(* Logix 5000 project; controller TFF vendor 1 type 14 code 107 rev 34.11; software revision 34.03; part 2 of 36 *)

        [3,10].HIHIAlarmONS := 1, [3,10].FeedPumpTag := 1, [3,10].Value := 4, [3,10].ValueHMI := 4, [3,10].PV := 20.567827, [3,10].HITimer.EN := 1, [3,10].HITimer.DN := 1, [3,10].HIHITimer.EN := 1, [3,10].HIHITimer.DN := 1, [3,10].EnableCfg := 1, [3,11].HIAlarm := 1, [3,11].HIHIAlarm := 1, [3,11].LOLODisable := 1, [3,11].LODisable := 1, [3,11].FeedPumpEnable := 1, [3,11].HIAlarmONS := 1, [3,11].HIHIAlarmONS := 1, [3,11].FeedPumpTag := 1, [3,11].Value := 4, [3,11].ValueHMI := 4, [3,11].PV := 25.7337, [3,11].HITimer.EN := 1, [3,11].HITimer.DN := 1, [3,11].HIHITimer.EN := 1, [3,11].HIHITimer.DN := 1, [3,11].EnableCfg := 1, [3,12].HIAlarm := 1, [3,12].HIHIAlarm := 1, [3,12].LOLODisable := 1, [3,12].LODisable := 1, [3,12].TransferPumpEnable := 1, [3,12].HIAlarmONS := 1, [3,12].HIHIAlarmONS := 1, [3,12].TransferPumpTag := 2, [3,12].Value := 4, [3,12].ValueHMI := 4, [3,12].PV := 28.0231, [3,12].HITimer.EN := 1, [3,12].HITimer.DN := 1, [3,12].HIHITimer.EN := 1, [3,12].HIHITimer.DN := 1, [3,12].EnableCfg := 1, [3,13].HIAlarm := 1, [3,13].HIHIAlarm := 1, [3,13].LOLODisable := 1, [3,13].LODisable := 1, [3,13].TransferPumpEnable := 1, [3,13].HIAlarmONS := 1, [3,13].HIHIAlarmONS := 1, [3,13].TransferPumpTag := 2, [3,13].Value := 4, [3,13].ValueHMI := 4, [3,13].PV := 21.08868, [3,13].HITimer.EN := 1, [3,13].HITimer.DN := 1, [3,13].HIHITimer.EN := 1, [3,13].HIHITimer.DN := 1, [3,13].EnableCfg := 1, [3,28].PV := -1.048729, [3,28].EnableCfg := 1,
        [3,29].HIAlarm := 1, [3,29].HIHIAlarm := 1, [3,29].HIAlarmONS := 1, [3,29].HIHIAlarmONS := 1, [3,29].Value := 4, [3,29].ValueHMI := 4, [3,29].PV := 100.96327, [3,29].HITimer.EN := 1, [3,29].HITimer.DN := 1, [3,29].HIHITimer.EN := 1, [3,29].HIHITimer.DN := 1, [3,29].EnableCfg := 1, [3,30].HIAlarm := 1, [3,30].HIHIAlarm := 1, [3,30].HIAlarmONS := 1, [3,30].HIHIAlarmONS := 1, [3,30].Value := 4, [3,30].ValueHMI := 4, [3,30].PV := 0.024414062, [3,30].HITimer.EN := 1, [3,30].HITimer.DN := 1, [3,30].HIHITimer.EN := 1, [3,30].HIHITimer.DN := 1, [3,30].EnableCfg := 1, [3,31].HIAlarm := 1, [3,31].HIHIAlarm := 1, [3,31].HIAlarmONS := 1, [3,31].HIHIAlarmONS := 1, [3,31].Value := 4, [3,31].ValueHMI := 4, [3,31].PV := 9.026997, [3,31].HITimer.EN := 1, [3,31].HITimer.DN := 1, [3,31].HIHITimer.EN := 1, [3,31].HIHITimer.DN := 1, [3,31].EnableCfg := 1, [3,40].LOLODisable := 1, [3,40].LODisable := 1, [3,40].FeedPumpEnable := 1, [3,40].TransferPumpEnable := 1, [3,40].FeedPumpTag := 1, [3,40].TransferPumpTag := 2, [3,40].PV := 48.590927, [3,40].EnableCfg := 1, [3,41].LOLODisable := 1, [3,41].LODisable := 1, [3,41].FeedPumpEnable := 1, [3,41].TransferPumpEnable := 1, [3,41].FeedPumpTag := 1, [3,41].TransferPumpTag := 2, [3,41].PV := 5830.911, [3,41].EnableCfg := 1, [3,42].LOLODisable := 1, [3,42].LODisable := 1, [3,42].FeedPumpEnable := 1, [3,42].FeedPumpTag := 1, [3,42].PV := 2468.1392, [3,42].EnableCfg := 1, [3,43].LOLODisable := 1, [3,43].LODisable := 1,
        [3,43].TransferPumpEnable := 1, [3,43].TransferPumpTag := 2, [3,43].PV := 3362.772, [3,43].EnableCfg := 1, [4,0].Override := 1, [4,0].LOLODisable := 1, [4,0].LODisable := 1, [4,0].LOLOAlarmONS := 1, [4,0].LOAlarmONS := 1, [4,0].HIAlarmONS := 1, [4,0].HIHIAlarmONS := 1, [4,0].HI := 100.0, [4,0].HIHI := 100.0, [4,0].PV := -2.4997964, [4,0].LOLOTimer.PRE := 2000, [4,0].LOLOTimerSP := 2, [4,0].LOTimer.PRE := 2000, [4,0].LOTimerSP := 2, [4,0].HITimer.PRE := 2000, [4,0].HITimerSP := 2, [4,0].HIHITimer.PRE := 2000, [4,0].HIHITimerSP := 2, [4,1].Override := 1, [4,1].LOLO := 20.0, [4,1].LO := 20.0, [4,1].HI := 50.0, [4,1].HIHI := 50.0, [4,1].PV := -12.498303, [4,1].LOLOTimer.PRE := 2000, [4,1].LOLOTimerSP := 2, [4,1].LOTimer.PRE := 2000, [4,1].LOTimerSP := 2, [4,1].HITimer.PRE := 2000, [4,1].HITimerSP := 2, [4,1].HIHITimer.PRE := 2000, [4,1].HIHITimerSP := 2, [4,1].EnableCfg := 1, [4,2].Override := 1, [4,2].LOLO := 20.0, [4,2].LO := 20.0, [4,2].HI := 100.0, [4,2].HIHI := 100.0, [4,2].PV := -24.996607, [4,2].LOLOTimer.PRE := 2000, [4,2].LOLOTimerSP := 2, [4,2].LOTimer.PRE := 2000, [4,2].LOTimerSP := 2, [4,2].HITimer.PRE := 2000, [4,2].HITimerSP := 2, [4,2].HIHITimer.PRE := 2000, [4,2].HIHITimerSP := 2, [4,2].EnableCfg := 1, [4,3].Override := 1, [4,3].LOLO := 5.0, [4,3].LO := 5.0, [4,3].HI := 14.0, [4,3].HIHI := 14.0, [4,3].PV := -3.499525, [4,3].LOLOTimer.PRE := 1000, [4,3].LOLOTimerSP := 1,
        [4,3].LOTimer.PRE := 5000, [4,3].LOTimerSP := 5, [4,3].HITimer.PRE := 5000, [4,3].HITimerSP := 5, [4,3].HIHITimer.PRE := 1000, [4,3].HIHITimerSP := 1, [4,3].EnableCfg := 1, [4,4].Override := 1, [4,4].HI := 100.0, [4,4].HIHI := 100.0, [4,4].PV := -24.996607, [4,4].LOLOTimer.PRE := 1000, [4,4].LOLOTimerSP := 1, [4,4].LOTimer.PRE := 5000, [4,4].LOTimerSP := 5, [4,4].HITimer.PRE := 5000, [4,4].HITimerSP := 5, [4,4].HIHITimer.PRE := 1000, [4,4].HIHITimerSP := 1, [4,4].EnableCfg := 1, [4,5].Override := 1, [4,5].LOLO := 2.0, [4,5].LO := 2.0, [4,5].HI := 3.0, [4,5].HIHI := 3.0, [4,5].PV := -0.7498982, [4,5].LOLOTimer.PRE := 2000, [4,5].LOLOTimerSP := 2, [4,5].LOTimer.PRE := 2000, [4,5].LOTimerSP := 2, [4,5].HITimer.PRE := 2000, [4,5].HITimerSP := 2, [4,5].HIHITimer.PRE := 2000, [4,5].HIHITimerSP := 2, [4,5].EnableCfg := 1, [4,6].Override := 1, [4,6].LOLO := 2.0, [4,6].LO := 2.0, [4,6].HI := 2.0, [4,6].HIHI := 2.0, [4,6].PV := -0.49993217, [4,6].LOLOTimer.PRE := 2000, [4,6].LOLOTimerSP := 2, [4,6].LOTimer.PRE := 2000, [4,6].LOTimerSP := 2, [4,6].HITimer.PRE := 2000, [4,6].HITimerSP := 2, [4,6].HIHITimer.PRE := 2000, [4,6].HIHITimerSP := 2, [4,6].EnableCfg := 1, [4,7].Override := 1, [4,7].LOLO := 20.0, [4,7].LO := 20.0, [4,7].HI := 100.0, [4,7].HIHI := 100.0, [4,7].PV := -24.996607, [4,7].LOLOTimer.PRE := 2000, [4,7].LOLOTimerSP := 2, [4,7].LOTimer.PRE := 2000, [4,7].LOTimerSP := 2,
        [4,7].HITimer.PRE := 2000, [4,7].HITimerSP := 2, [4,7].HIHITimer.PRE := 2000, [4,7].HIHITimerSP := 2, [4,7].EnableCfg := 1, [4,8].Override := 1, [4,8].HI := 14.0, [4,8].HIHI := 14.0, [4,8].PV := -3.499525, [4,8].LOLOTimer.PRE := 1000, [4,8].LOLOTimerSP := 1, [4,8].LOTimer.PRE := 5000, [4,8].LOTimerSP := 5, [4,8].HITimer.PRE := 5000, [4,8].HITimerSP := 5, [4,8].HIHITimer.PRE := 1000, [4,8].HIHITimerSP := 1, [4,8].EnableCfg := 1, [4,9].Override := 1, [4,9].LOLODisable := 1, [4,9].LODisable := 1, [4,9].FeedPumpEnable := 1, [4,9].TransferPumpEnable := 1, [4,9].FeedPumpTag := 1, [4,9].TransferPumpTag := 2, [4,9].HI := 6.0, [4,9].HIHI := 6.0, [4,9].PV := -1.4998856, [4,9].LOLOTimer.PRE := 2000, [4,9].LOLOTimerSP := 2, [4,9].LOTimer.PRE := 2000, [4,9].LOTimerSP := 2, [4,9].HITimer.PRE := 2000, [4,9].HITimerSP := 2, [4,9].HIHITimer.PRE := 2000, [4,9].HIHITimerSP := 2, [4,9].EnableCfg := 1, [4,10].Override := 1, [4,10].LOLODisable := 1, [4,10].LODisable := 1, [4,10].FeedPumpEnable := 1, [4,10].FeedPumpTag := 1, [4,10].HI := 22.0, [4,10].HIHI := 22.0, [4,10].LOLOTimer.PRE := 2000, [4,10].LOLOTimerSP := 2, [4,10].LOTimer.PRE := 2000, [4,10].LOTimerSP := 2, [4,10].HITimer.PRE := 2000, [4,10].HITimerSP := 2, [4,10].HIHITimer.PRE := 2000, [4,10].HIHITimerSP := 2, [4,10].EnableCfg := 1, [4,11].Override := 1, [4,11].LOLODisable := 1, [4,11].LODisable := 1, [4,11].FeedPumpEnable := 1, [4,11].FeedPumpTag := 1, [4,11].HI := 6.0, [4,11].HIHI := 6.0,
        [4,11].PV := -1.4998856, [4,11].LOLOTimer.PRE := 2000, [4,11].LOLOTimerSP := 2, [4,11].LOTimer.PRE := 2000, [4,11].LOTimerSP := 2, [4,11].HITimer.PRE := 2000, [4,11].HITimerSP := 2, [4,11].HIHITimer.PRE := 2000, [4,11].HIHITimerSP := 2, [4,11].EnableCfg := 1, [4,12].Override := 1, [4,12].LOLODisable := 1, [4,12].LODisable := 1, [4,12].TransferPumpEnable := 1, [4,12].TransferPumpTag := 2, [4,12].HI := 22.0, [4,12].HIHI := 22.0, [4,12].LOLOTimer.PRE := 2000, [4,12].LOLOTimerSP := 2, [4,12].LOTimer.PRE := 2000, [4,12].LOTimerSP := 2, [4,12].HITimer.PRE := 2000, [4,12].HITimerSP := 2, [4,12].HIHITimer.PRE := 2000, [4,12].HIHITimerSP := 2, [4,12].EnableCfg := 1, [4,13].Override := 1, [4,13].LOLODisable := 1, [4,13].LODisable := 1, [4,13].TransferPumpEnable := 1, [4,13].TransferPumpTag := 2, [4,13].HI := 6.0, [4,13].HIHI := 6.0, [4,13].PV := -1.4998856, [4,13].LOLOTimer.PRE := 2000, [4,13].LOLOTimerSP := 2, [4,13].LOTimer.PRE := 2000, [4,13].LOTimerSP := 2, [4,13].HITimer.PRE := 2000, [4,13].HITimerSP := 2, [4,13].HIHITimer.PRE := 2000, [4,13].HIHITimerSP := 2, [4,13].EnableCfg := 1, [4,14].Override := 1, [4,14].HI := 14.0, [4,14].HIHI := 14.0, [4,14].LOLOTimer.PRE := 1000, [4,14].LOLOTimerSP := 1, [4,14].LOTimer.PRE := 5000, [4,14].LOTimerSP := 5, [4,14].HITimer.PRE := 5000, [4,14].HITimerSP := 5, [4,14].HIHITimer.PRE := 1000, [4,14].HIHITimerSP := 1, [4,15].Override := 1, [4,15].HI := 2.0, [4,15].HIHI := 2.0, [4,15].PV := -0.49993217, [4,15].LOLOTimer.PRE := 2000, [4,15].LOLOTimerSP := 2,
        [4,15].LOTimer.PRE := 2000, [4,15].LOTimerSP := 2, [4,15].HITimer.PRE := 2000, [4,15].HITimerSP := 2, [4,15].HIHITimer.PRE := 2000, [4,15].HIHITimerSP := 2, [4,16].Override := 1, [4,16].HI := 2.0, [4,16].HIHI := 2.0, [4,16].PV := -0.49993217, [4,16].LOLOTimer.PRE := 2000, [4,16].LOLOTimerSP := 2, [4,16].LOTimer.PRE := 2000, [4,16].LOTimerSP := 2, [4,16].HITimer.PRE := 2000, [4,16].HITimerSP := 2, [4,16].HIHITimer.PRE := 2000, [4,16].HIHITimerSP := 2, [4,17].Override := 1, [4,17].LOLODisable := 1, [4,17].LODisable := 1, [4,17].FeedPumpEnable := 1, [4,17].TransferPumpEnable := 1, [4,17].FeedPumpTag := 1, [4,17].TransferPumpTag := 2, [4,17].LOLO := -1.0, [4,17].LO := -1.0, [4,17].HI := 5.0, [4,17].HIHI := 5.0, [4,17].PV := -2.4997964, [4,17].LOLOTimer.PRE := 2000, [4,17].LOLOTimerSP := 2, [4,17].LOTimer.PRE := 2000, [4,17].LOTimerSP := 2, [4,17].HITimer.PRE := 2000, [4,17].HITimerSP := 2, [4,17].HIHITimer.PRE := 2000, [4,17].HIHITimerSP := 2, [4,18].Override := 1, [4,18].LOLODisable := 1, [4,18].LODisable := 1, [4,18].FeedPumpEnable := 1, [4,18].FeedPumpTag := 1, [4,18].LOLO := -1.0, [4,18].LO := -1.0, [4,18].HI := 5.0, [4,18].HIHI := 5.0, [4,18].PV := -2.4997964, [4,18].LOLOTimer.PRE := 2000, [4,18].LOLOTimerSP := 2, [4,18].LOTimer.PRE := 2000, [4,18].LOTimerSP := 2, [4,18].HITimer.PRE := 2000, [4,18].HITimerSP := 2, [4,18].HIHITimer.PRE := 2000, [4,18].HIHITimerSP := 2, [4,19].Override := 1, [4,19].LOLODisable := 1, [4,19].LODisable := 1, [4,19].TransferPumpEnable := 1,
        [4,19].TransferPumpTag := 2, [4,19].LOLO := -1.0, [4,19].LO := -1.0, [4,19].HI := 5.0, [4,19].HIHI := 5.0, [4,19].PV := -2.4997964, [4,19].LOLOTimer.PRE := 2000, [4,19].LOLOTimerSP := 2, [4,19].LOTimer.PRE := 2000, [4,19].LOTimerSP := 2, [4,19].HITimer.PRE := 2000, [4,19].HITimerSP := 2, [4,19].HIHITimer.PRE := 2000, [4,19].HIHITimerSP := 2, [4,20].Override := 1, [4,20].HI := 100.0, [4,20].HIHI := 100.0, [4,20].PV := 100.0, [4,20].LOLOTimerSP := 2, [4,20].LOTimerSP := 2, [4,20].HITimer.EN := 1, [4,20].HITimer.DN := 1, [4,20].HITimerSP := 2, [4,20].HIHITimer.EN := 1, [4,20].HIHITimer.DN := 1, [4,20].HIHITimerSP := 2, [4,21].Override := 1, [4,21].HI := 100.0, [4,21].HIHI := 100.0, [4,21].LOLOTimerSP := 2, [4,21].LOTimerSP := 2, [4,21].HITimerSP := 2, [4,21].HIHITimerSP := 2, [4,22].Override := 1, [4,22].PV := 0.50476843, [4,23].Override := 1, [4,23].PV := 0.11619745, [4,24].Override := 1, [4,24].PV := 0.16, [4,25].Override := 1, [4,25].PV := -0.3333333, [4,26].Override := 1, [4,26].PV := 63.88032, [4,27].Override := 1, [4,27].PV := -37.40687, [4,28].Override := 1, [4,28].HI := 100.0, [4,28].HIHI := 100.0, [4,28].PV := 22.8542, [4,28].LOLOTimer.PRE := 2000, [4,28].LOLOTimerSP := 2, [4,28].LOTimer.PRE := 2000, [4,28].LOTimerSP := 2, [4,28].HITimer.PRE := 2000, [4,28].HITimerSP := 2, [4,28].HIHITimer.PRE := 2000, [4,28].HIHITimerSP := 2, [4,28].EnableCfg := 1, [4,29].Override := 1, [4,29].HI := 100.0,
        [4,29].HIHI := 100.0, [4,29].PV := 21.877623, [4,29].LOLOTimer.PRE := 2000, [4,29].LOLOTimerSP := 2, [4,29].LOTimer.PRE := 2000, [4,29].LOTimerSP := 2, [4,29].HITimer.PRE := 2000, [4,29].HITimerSP := 2, [4,29].HIHITimer.PRE := 2000, [4,29].HIHITimerSP := 2, [4,29].EnableCfg := 1, [4,30].Override := 1, [4,30].HI := 100.0, [4,30].HIHI := 100.0, [4,30].PV := 21.877623, [4,30].LOLOTimer.PRE := 2000, [4,30].LOLOTimerSP := 2, [4,30].LOTimer.PRE := 2000, [4,30].LOTimerSP := 2, [4,30].HITimer.PRE := 2000, [4,30].HITimerSP := 2, [4,30].HIHITimer.PRE := 2000, [4,30].HIHITimerSP := 2, [4,30].EnableCfg := 1, [4,31].Override := 1, [4,31].HI := 100.0, [4,31].HIHI := 100.0, [4,31].PV := 21.877623, [4,31].LOLOTimer.PRE := 2000, [4,31].LOLOTimerSP := 2, [4,31].LOTimer.PRE := 2000, [4,31].LOTimerSP := 2, [4,31].HITimer.PRE := 2000, [4,31].HITimerSP := 2, [4,31].HIHITimer.PRE := 2000, [4,31].HIHITimerSP := 2, [4,31].EnableCfg := 1, [4,32].Override := 1, [4,32].PV := 0.1837702, [4,33].Override := 1, [4,33].PV := -0.6615715, [4,34].Override := 1, [4,34].PV := 0.6615715, [4,35].Override := 1, [4,35].PV := 222.0, [4,36].Override := 1, [4,37].Override := 1, [4,37].PV := -0.03181506, [4,38].Override := 1, [4,39].Override := 1, [4,40].Override := 1, [4,40].LOLODisable := 1, [4,40].LODisable := 1, [4,40].FeedPumpEnable := 1, [4,40].TransferPumpEnable := 1, [4,40].FeedPumpTag := 1, [4,40].TransferPumpTag := 2, [4,40].HI := 44.0, [4,40].HIHI := 44.0, [4,40].LOLOTimer.PRE := 2000,
        [4,40].LOLOTimerSP := 2, [4,40].LOTimer.PRE := 2000, [4,40].LOTimerSP := 2, [4,40].HITimer.PRE := 2000, [4,40].HITimerSP := 2, [4,40].HIHITimer.PRE := 2000, [4,40].HIHITimerSP := 2, [4,40].EnableCfg := 1, [4,41].Override := 1, [4,41].LOLODisable := 1, [4,41].LODisable := 1, [4,41].FeedPumpEnable := 1, [4,41].TransferPumpEnable := 1, [4,41].FeedPumpTag := 1, [4,41].TransferPumpTag := 2, [4,41].HI := 9999.0, [4,41].HIHI := 9999.0, [4,41].LOLOTimer.PRE := 2000, [4,41].LOLOTimerSP := 2, [4,41].LOTimer.PRE := 2000, [4,41].LOTimerSP := 2, [4,41].HITimer.PRE := 2000, [4,41].HITimerSP := 2, [4,41].HIHITimer.PRE := 2000, [4,41].HIHITimerSP := 2, [4,41].EnableCfg := 1, [4,42].Override := 1, [4,42].LOLODisable := 1, [4,42].LODisable := 1, [4,42].FeedPumpEnable := 1, [4,42].FeedPumpTag := 1, [4,42].HI := 9999.0, [4,42].HIHI := 9999.0, [4,42].LOLOTimer.PRE := 2000, [4,42].LOLOTimerSP := 2, [4,42].LOTimer.PRE := 2000, [4,42].LOTimerSP := 2, [4,42].HITimer.PRE := 2000, [4,42].HITimerSP := 2, [4,42].HIHITimer.PRE := 2000, [4,42].HIHITimerSP := 2, [4,42].EnableCfg := 1, [4,43].Override := 1, [4,43].LOLODisable := 1, [4,43].LODisable := 1, [4,43].TransferPumpEnable := 1, [4,43].TransferPumpTag := 2, [4,43].HI := 9999.0, [4,43].HIHI := 9999.0, [4,43].LOLOTimer.PRE := 2000, [4,43].LOLOTimerSP := 2, [4,43].LOTimer.PRE := 2000, [4,43].LOTimerSP := 2, [4,43].HITimer.PRE := 2000, [4,43].HITimerSP := 2, [4,43].HIHITimer.PRE := 2000, [4,43].HIHITimerSP := 2, [4,43].EnableCfg := 1, [4,44].Override := 1, [4,44].HI := 99999.0,
        [4,44].HIHI := 99999.0, [4,44].LOLOTimerSP := 2, [4,44].LOTimerSP := 2, [4,44].HITimerSP := 2, [4,44].HIHITimerSP := 2, [4,45].Override := 1, [4,45].Disable := 1, [4,45].LOLODisable := 1, [4,45].LODisable := 1, [4,45].FeedPumpEnable := 1, [4,45].TransferPumpEnable := 1, [4,45].FeedPumpTag := 1, [4,45].TransferPumpTag := 2, [4,45].LOLO := -1.0, [4,45].LO := -1.0, [4,45].HI := 5.0, [4,45].HIHI := 5.0, [4,45].LOLOTimer.PRE := 2000, [4,45].LOLOTimerSP := 2, [4,45].LOTimer.PRE := 2000, [4,45].LOTimerSP := 2, [4,45].HITimer.PRE := 2000, [4,45].HITimerSP := 2, [4,45].HIHITimer.PRE := 2000, [4,45].HIHITimerSP := 2, [4,46].Override := 1, [4,47].Override := 1, [4,48].Override := 1, [4,49].Override := 1, [5,0].Override := 1, [5,0].LOLODisable := 1, [5,0].LODisable := 1, [5,0].LOLOAlarmONS := 1, [5,0].LOAlarmONS := 1, [5,0].HIAlarmONS := 1, [5,0].HIHIAlarmONS := 1, [5,0].HI := 100.0, [5,0].HIHI := 100.0, [5,0].PV := -2.4997964, [5,0].LOLOTimer.PRE := 2000, [5,0].LOLOTimerSP := 2, [5,0].LOTimer.PRE := 2000, [5,0].LOTimerSP := 2, [5,0].HITimer.PRE := 2000, [5,0].HITimerSP := 2, [5,0].HIHITimer.PRE := 2000, [5,0].HIHITimerSP := 2, [5,1].Override := 1, [5,1].LOLODisable := 1, [5,1].LODisable := 1, [5,1].HI := 50.0, [5,1].HIHI := 50.0, [5,1].PV := -6.249152, [5,1].LOLOTimer.PRE := 2000, [5,1].LOLOTimerSP := 2, [5,1].LOTimer.PRE := 2000, [5,1].LOTimerSP := 2, [5,1].HITimer.PRE := 2000, [5,1].HITimerSP := 2, [5,1].HIHITimer.PRE := 2000,
        [5,1].HIHITimerSP := 2, [5,1].EnableCfg := 1, [5,2].Override := 1, [5,2].LOLODisable := 1, [5,2].LODisable := 1, [5,2].HI := 100.0, [5,2].HIHI := 100.0, [5,2].PV := -2.4997966, [5,2].LOLOTimer.PRE := 2000, [5,2].LOLOTimerSP := 2, [5,2].LOTimer.PRE := 2000, [5,2].LOTimerSP := 2, [5,2].HITimer.PRE := 2000, [5,2].HITimerSP := 2, [5,2].HIHITimer.PRE := 2000, [5,2].HIHITimerSP := 2, [5,2].EnableCfg := 1, [5,3].Override := 1, [5,3].LOLODisable := 1, [5,3].LODisable := 1, [5,3].HI := 14.0, [5,3].HIHI := 14.0, [5,3].PV := -6.249152, [5,3].LOLOTimer.PRE := 1000, [5,3].LOLOTimerSP := 1, [5,3].LOTimer.PRE := 5000, [5,3].LOTimerSP := 5, [5,3].HITimer.PRE := 5000, [5,3].HITimerSP := 5, [5,3].HIHITimer.PRE := 1000, [5,3].HIHITimerSP := 1, [5,3].EnableCfg := 1, [5,4].Override := 1, [5,4].HI := 100.0, [5,4].HIHI := 100.0, [5,4].PV := -37.49491, [5,4].LOLOTimer.PRE := 1000, [5,4].LOLOTimerSP := 1, [5,4].LOTimer.PRE := 5000, [5,4].LOTimerSP := 5, [5,4].HITimer.PRE := 5000, [5,4].HITimerSP := 5, [5,4].HIHITimer.PRE := 1000, [5,4].HIHITimerSP := 1, [5,4].EnableCfg := 1, [5,5].Override := 1, [5,5].HI := 2.0, [5,5].HIHI := 2.0, [5,5].PV := -37.49491, [5,5].LOLOTimer.PRE := 2000, [5,5].LOLOTimerSP := 2, [5,5].LOTimer.PRE := 2000, [5,5].LOTimerSP := 2, [5,5].HITimer.PRE := 2000, [5,5].HITimerSP := 2, [5,5].HIHITimer.PRE := 2000, [5,5].HIHITimerSP := 2, [5,5].EnableCfg := 1, [5,6].Override := 1, [5,6].LOLODisable := 1,
        [5,6].LODisable := 1, [5,6].HI := 2.0, [5,6].HIHI := 2.0, [5,6].PV := -2.4997966, [5,6].LOLOTimer.PRE := 2000, [5,6].LOLOTimerSP := 2, [5,6].LOTimer.PRE := 2000, [5,6].LOTimerSP := 2, [5,6].HITimer.PRE := 2000, [5,6].HITimerSP := 2, [5,6].HIHITimer.PRE := 2000, [5,6].HIHITimerSP := 2, [5,6].EnableCfg := 1, [5,7].Override := 1, [5,7].LOLODisable := 1, [5,7].LODisable := 1, [5,7].HI := 100.0, [5,7].HIHI := 100.0, [5,7].PV := -2.4997966, [5,7].LOLOTimer.PRE := 2000, [5,7].LOLOTimerSP := 2, [5,7].LOTimer.PRE := 2000, [5,7].LOTimerSP := 2, [5,7].HITimer.PRE := 2000, [5,7].HITimerSP := 2, [5,7].HIHITimer.PRE := 2000, [5,7].HIHITimerSP := 2, [5,7].EnableCfg := 1, [5,8].Override := 1, [5,8].HI := 14.0, [5,8].HIHI := 14.0, [5,8].PV := -49.993217, [5,8].LOLOTimer.PRE := 1000, [5,8].LOLOTimerSP := 1, [5,8].LOTimer.PRE := 5000, [5,8].LOTimerSP := 5, [5,8].HITimer.PRE := 5000, [5,8].HITimerSP := 5, [5,8].HIHITimer.PRE := 1000, [5,8].HIHITimerSP := 1, [5,8].EnableCfg := 1, [5,9].Override := 1, [5,9].LOLODisable := 1, [5,9].LODisable := 1, [5,9].FeedPumpEnable := 1, [5,9].TransferPumpEnable := 1, [5,9].FeedPumpTag := 1, [5,9].TransferPumpTag := 2, [5,9].HI := 6.0, [5,9].HIHI := 6.0, [5,9].PV := -3.499733, [5,9].LOLOTimer.PRE := 2000, [5,9].LOLOTimerSP := 2, [5,9].LOTimer.PRE := 2000, [5,9].LOTimerSP := 2, [5,9].HITimer.PRE := 2000, [5,9].HITimerSP := 2, [5,9].HIHITimer.PRE := 2000, [5,9].HIHITimerSP := 2, [5,9].EnableCfg := 1,
        [5,10].Override := 1, [5,10].LOLODisable := 1, [5,10].LODisable := 1, [5,10].FeedPumpEnable := 1, [5,10].FeedPumpTag := 1, [5,10].HI := 22.0, [5,10].HIHI := 22.0, [5,10].LOLOTimer.PRE := 2000, [5,10].LOLOTimerSP := 2, [5,10].LOTimer.PRE := 2000, [5,10].LOTimerSP := 2, [5,10].HITimer.PRE := 2000, [5,10].HITimerSP := 2, [5,10].HIHITimer.PRE := 2000, [5,10].HIHITimerSP := 2, [5,10].EnableCfg := 1, [5,11].Override := 1, [5,11].LOLODisable := 1, [5,11].LODisable := 1, [5,11].FeedPumpEnable := 1, [5,11].FeedPumpTag := 1, [5,11].HI := 6.0, [5,11].HIHI := 6.0, [5,11].PV := -49.996185, [5,11].LOLOTimer.PRE := 2000, [5,11].LOLOTimerSP := 2, [5,11].LOTimer.PRE := 2000, [5,11].LOTimerSP := 2, [5,11].HITimer.PRE := 2000, [5,11].HITimerSP := 2, [5,11].HIHITimer.PRE := 2000, [5,11].HIHITimerSP := 2, [5,11].EnableCfg := 1, [5,12].Override := 1, [5,12].LOLODisable := 1, [5,12].LODisable := 1, [5,12].TransferPumpEnable := 1, [5,12].TransferPumpTag := 2, [5,12].HI := 22.0, [5,12].HIHI := 22.0, [5,12].LOLOTimer.PRE := 2000, [5,12].LOLOTimerSP := 2, [5,12].LOTimer.PRE := 2000, [5,12].LOTimerSP := 2, [5,12].HITimer.PRE := 2000, [5,12].HITimerSP := 2, [5,12].HIHITimer.PRE := 2000, [5,12].HIHITimerSP := 2, [5,12].EnableCfg := 1, [5,13].Override := 1, [5,13].LOLODisable := 1, [5,13].LODisable := 1, [5,13].TransferPumpEnable := 1, [5,13].TransferPumpTag := 2, [5,13].HI := 6.0, [5,13].HIHI := 6.0, [5,13].PV := -24.998093, [5,13].LOLOTimer.PRE := 2000, [5,13].LOLOTimerSP := 2, [5,13].LOTimer.PRE := 2000,
        [5,13].LOTimerSP := 2, [5,13].HITimer.PRE := 2000, [5,13].HITimerSP := 2, [5,13].HIHITimer.PRE := 2000, [5,13].HIHITimerSP := 2, [5,13].EnableCfg := 1, [5,14].Override := 1, [5,14].HI := 14.0, [5,14].HIHI := 14.0, [5,14].LOLOTimer.PRE := 1000, [5,14].LOLOTimerSP := 1, [5,14].LOTimer.PRE := 5000, [5,14].LOTimerSP := 5, [5,14].HITimer.PRE := 5000, [5,14].HITimerSP := 5, [5,14].HIHITimer.PRE := 1000, [5,14].HIHITimerSP := 1, [5,15].Override := 1, [5,15].HI := 2.0, [5,15].HIHI := 2.0, [5,15].PV := -0.49993217, [5,15].LOLOTimer.PRE := 2000, [5,15].LOLOTimerSP := 2, [5,15].LOTimer.PRE := 2000, [5,15].LOTimerSP := 2, [5,15].HITimer.PRE := 2000, [5,15].HITimerSP := 2, [5,15].HIHITimer.PRE := 2000, [5,15].HIHITimerSP := 2, [5,16].Override := 1, [5,16].HI := 2.0, [5,16].HIHI := 2.0, [5,16].PV := -0.49993217, [5,16].LOLOTimer.PRE := 2000, [5,16].LOLOTimerSP := 2, [5,16].LOTimer.PRE := 2000, [5,16].LOTimerSP := 2, [5,16].HITimer.PRE := 2000, [5,16].HITimerSP := 2, [5,16].HIHITimer.PRE := 2000, [5,16].HIHITimerSP := 2, [5,17].Override := 1, [5,17].LOLODisable := 1, [5,17].LODisable := 1, [5,17].FeedPumpEnable := 1, [5,17].TransferPumpEnable := 1, [5,17].FeedPumpTag := 1, [5,17].TransferPumpTag := 2, [5,17].LOLO := -1.0, [5,17].LO := -1.0, [5,17].HI := 5.0, [5,17].HIHI := 5.0, [5,17].PV := -2.4997964, [5,17].LOLOTimer.PRE := 2000, [5,17].LOLOTimerSP := 2, [5,17].LOTimer.PRE := 2000, [5,17].LOTimerSP := 2, [5,17].HITimer.PRE := 2000, [5,17].HITimerSP := 2, [5,17].HIHITimer.PRE := 2000,
        [5,17].HIHITimerSP := 2, [5,18].Override := 1, [5,18].LOLODisable := 1, [5,18].LODisable := 1, [5,18].FeedPumpEnable := 1, [5,18].FeedPumpTag := 1, [5,18].LOLO := -1.0, [5,18].LO := -1.0, [5,18].HI := 5.0, [5,18].HIHI := 5.0, [5,18].PV := -2.4997964, [5,18].LOLOTimer.PRE := 2000, [5,18].LOLOTimerSP := 2, [5,18].LOTimer.PRE := 2000, [5,18].LOTimerSP := 2, [5,18].HITimer.PRE := 2000, [5,18].HITimerSP := 2, [5,18].HIHITimer.PRE := 2000, [5,18].HIHITimerSP := 2, [5,19].Override := 1, [5,19].LOLODisable := 1, [5,19].LODisable := 1, [5,19].TransferPumpEnable := 1, [5,19].TransferPumpTag := 2, [5,19].LOLO := -1.0, [5,19].LO := -1.0, [5,19].HI := 5.0, [5,19].HIHI := 5.0, [5,19].PV := -2.4997964, [5,19].LOLOTimer.PRE := 2000, [5,19].LOLOTimerSP := 2, [5,19].LOTimer.PRE := 2000, [5,19].LOTimerSP := 2, [5,19].HITimer.PRE := 2000, [5,19].HITimerSP := 2, [5,19].HIHITimer.PRE := 2000, [5,19].HIHITimerSP := 2, [5,20].Override := 1, [5,20].HI := 100.0, [5,20].HIHI := 100.0, [5,20].PV := 100.0, [5,20].LOLOTimerSP := 2, [5,20].LOTimerSP := 2, [5,20].HITimer.EN := 1, [5,20].HITimer.DN := 1, [5,20].HITimerSP := 2, [5,20].HIHITimer.EN := 1, [5,20].HIHITimer.DN := 1, [5,20].HIHITimerSP := 2, [5,21].Override := 1, [5,21].HI := 100.0, [5,21].HIHI := 100.0, [5,21].LOLOTimerSP := 2, [5,21].LOTimerSP := 2, [5,21].HITimerSP := 2, [5,21].HIHITimerSP := 2, [5,22].Override := 1, [5,22].PV := 0.50476843, [5,23].Override := 1, [5,23].PV := 0.11619745,
        [5,24].Override := 1, [5,24].PV := 0.16, [5,25].Override := 1, [5,25].PV := -0.3333333, [5,26].Override := 1, [5,26].PV := 63.88032, [5,27].Override := 1, [5,27].PV := -37.40687, [5,28].Override := 1, [5,28].HI := 100.0, [5,28].HIHI := 100.0, [5,28].PV := -24.998093, [5,28].LOLOTimer.PRE := 2000, [5,28].LOLOTimerSP := 2, [5,28].LOTimer.PRE := 2000, [5,28].LOTimerSP := 2, [5,28].HITimer.PRE := 2000, [5,28].HITimerSP := 2, [5,28].HIHITimer.PRE := 2000, [5,28].HIHITimerSP := 2, [5,28].EnableCfg := 1, [5,29].Override := 1, [5,29].HI := 100.0, [5,29].HIHI := 100.0, [5,29].PV := -24.998093, [5,29].LOLOTimer.PRE := 2000, [5,29].LOLOTimerSP := 2, [5,29].LOTimer.PRE := 2000, [5,29].LOTimerSP := 2, [5,29].HITimer.PRE := 2000, [5,29].HITimerSP := 2, [5,29].HIHITimer.PRE := 2000, [5,29].HIHITimerSP := 2, [5,29].EnableCfg := 1, [5,30].Override := 1, [5,30].HI := 100.0, [5,30].HIHI := 100.0, [5,30].PV := -24.998093, [5,30].LOLOTimer.PRE := 2000, [5,30].LOLOTimerSP := 2, [5,30].LOTimer.PRE := 2000, [5,30].LOTimerSP := 2, [5,30].HITimer.PRE := 2000, [5,30].HITimerSP := 2, [5,30].HIHITimer.PRE := 2000, [5,30].HIHITimerSP := 2, [5,30].EnableCfg := 1, [5,31].Override := 1, [5,31].HI := 100.0, [5,31].HIHI := 100.0, [5,31].PV := -24.998093, [5,31].LOLOTimer.PRE := 2000, [5,31].LOLOTimerSP := 2, [5,31].LOTimer.PRE := 2000, [5,31].LOTimerSP := 2, [5,31].HITimer.PRE := 2000, [5,31].HITimerSP := 2, [5,31].HIHITimer.PRE := 2000, [5,31].HIHITimerSP := 2, [5,31].EnableCfg := 1,
        [5,32].Override := 1, [5,32].PV := 0.1837702, [5,33].Override := 1, [5,33].PV := -0.6615715, [5,34].Override := 1, [5,34].PV := 0.6615715, [5,35].Override := 1, [5,35].PV := 222.0, [5,36].Override := 1, [5,37].Override := 1, [5,37].PV := -0.03181506, [5,38].Override := 1, [5,39].Override := 1, [5,40].Override := 1, [5,40].LOLODisable := 1, [5,40].LODisable := 1, [5,40].FeedPumpEnable := 1, [5,40].TransferPumpEnable := 1, [5,40].FeedPumpTag := 1, [5,40].TransferPumpTag := 2, [5,40].HI := 44.0, [5,40].HIHI := 44.0, [5,40].LOLOTimer.PRE := 2000, [5,40].LOLOTimerSP := 2, [5,40].LOTimer.PRE := 2000, [5,40].LOTimerSP := 2, [5,40].HITimer.PRE := 2000, [5,40].HITimerSP := 2, [5,40].HIHITimer.PRE := 2000, [5,40].HIHITimerSP := 2, [5,40].EnableCfg := 1, [5,41].Override := 1, [5,41].LOLODisable := 1, [5,41].LODisable := 1, [5,41].FeedPumpEnable := 1, [5,41].TransferPumpEnable := 1, [5,41].FeedPumpTag := 1, [5,41].TransferPumpTag := 2, [5,41].HI := 9999.0, [5,41].HIHI := 9999.0, [5,41].LOLOTimer.PRE := 2000, [5,41].LOLOTimerSP := 2, [5,41].LOTimer.PRE := 2000, [5,41].LOTimerSP := 2, [5,41].HITimer.PRE := 2000, [5,41].HITimerSP := 2, [5,41].HIHITimer.PRE := 2000, [5,41].HIHITimerSP := 2, [5,41].EnableCfg := 1, [5,42].Override := 1, [5,42].LOLODisable := 1, [5,42].LODisable := 1, [5,42].FeedPumpEnable := 1, [5,42].FeedPumpTag := 1, [5,42].HI := 9999.0, [5,42].HIHI := 9999.0, [5,42].LOLOTimer.PRE := 2000, [5,42].LOLOTimerSP := 2, [5,42].LOTimer.PRE := 2000, [5,42].LOTimerSP := 2,
        [5,42].HITimer.PRE := 2000, [5,42].HITimerSP := 2, [5,42].HIHITimer.PRE := 2000, [5,42].HIHITimerSP := 2, [5,42].EnableCfg := 1, [5,43].Override := 1, [5,43].LOLODisable := 1, [5,43].LODisable := 1, [5,43].TransferPumpEnable := 1, [5,43].TransferPumpTag := 2, [5,43].HI := 9999.0, [5,43].HIHI := 9999.0, [5,43].LOLOTimer.PRE := 2000, [5,43].LOLOTimerSP := 2, [5,43].LOTimer.PRE := 2000, [5,43].LOTimerSP := 2, [5,43].HITimer.PRE := 2000, [5,43].HITimerSP := 2, [5,43].HIHITimer.PRE := 2000, [5,43].HIHITimerSP := 2, [5,43].EnableCfg := 1, [5,44].Override := 1, [5,44].HI := 99999.0, [5,44].HIHI := 99999.0, [5,44].LOLOTimerSP := 2, [5,44].LOTimerSP := 2, [5,44].HITimerSP := 2, [5,44].HIHITimerSP := 2, [5,45].Override := 1, [5,45].Disable := 1, [5,45].LOLODisable := 1, [5,45].LODisable := 1, [5,45].FeedPumpEnable := 1, [5,45].TransferPumpEnable := 1, [5,45].FeedPumpTag := 1, [5,45].TransferPumpTag := 2, [5,45].LOLO := -1.0, [5,45].LO := -1.0, [5,45].HI := 5.0, [5,45].HIHI := 5.0, [5,45].LOLOTimer.PRE := 2000, [5,45].LOLOTimerSP := 2, [5,45].LOTimer.PRE := 2000, [5,45].LOTimerSP := 2, [5,45].HITimer.PRE := 2000, [5,45].HITimerSP := 2, [5,45].HIHITimer.PRE := 2000, [5,45].HIHITimerSP := 2, [5,46].Override := 1, [5,47].Override := 1, [5,48].Override := 1, [5,49].Override := 1);
   AlarmControl : AlarmControl := (AlarmLow := 1, AlarmLowUnack := 1, LowHMI := 1, LowUnackHMI := 1, Horn := 1, Current := 1, FlashTimer.PRE := 500, FlashTimer.ACC := 251, FlashTimer.EN := 1, FlashTimer.TT := 1, AckTimer.PRE := 3000, EnableAllTimer.PRE := 3000, DisableAllTimer.PRE := 3000, HornAddress := 1, EnableAllAnaSigTimer.PRE := 3000, DisableAllAnaSigTimer.PRE := 3000, ESAckTimer.PRE := 3000);   // Alarm Control
        .FlashTimer.DN   // Alarm Control
   AlarmDeviation : AlarmDeviation[20] := ([0].Override := 1, [0].Disable := 1, [0].HIAlarmONS := 1, [0].HIHIAlarmONS := 1, [0].HI := 40.0, [0].HIHI := 53.0, [0].LOLOLim := 31.33333, [0].LOLim := 39.99999, [0].HILim := 93.33332, [0].HIHILim := 102.0, [0].HITimer.PRE := 30000, [0].HIHITimer.PRE := 30000, [1].Override := 1, [1].Disable := 1, [1].HI := 100.0, [1].HIHI := 100.0, [1].HILim := 20.0, [1].HIHILim := 20.0, [1].HITimer.PRE := 2000, [1].HITimerSP := 2, [1].HIHITimer.PRE := 2000, [1].HIHITImerSP := 2, [1].EnableCfg := 1, [2].Override := 1, [2].Disable := 1, [2].HI := 100.0, [2].HIHI := 100.0, [2].HILim := 103.18, [2].HIHILim := 103.18, [2].HITimer.PRE := 2000, [2].HITimerSP := 2, [2].HIHITimer.PRE := 2000, [2].HIHITImerSP := 2, [2].EnableCfg := 1, [3].Override := 1, [3].Disable := 1, [3].HI := 100.0, [3].HIHI := 100.0, [3].HILim := 12.0, [3].HIHILim := 12.0, [3].HITimer.PRE := 5000, [3].HITimerSP := 5, [3].HIHITimer.PRE := 5000, [3].HIHITImerSP := 5, [3].EnableCfg := 1, [4].Override := 1, [4].Disable := 1, [4].HI := 100.0, [4].HIHI := 100.0, [4].HITimer.PRE := 2000, [4].HITimerSP := 2, [4].HIHITimer.PRE := 2000, [4].HIHITImerSP := 2, [5].Override := 1, [5].Disable := 1, [5].HI := 100.0, [5].HIHI := 100.0, [5].EnableCfg := 1, [6].Override := 1, [6].Disable := 1,
        [6].HI := 100.0, [6].HIHI := 100.0, [6].HITimer.PRE := 2000, [6].HITimerSP := 2, [6].HIHITimer.PRE := 2000, [6].HIHITImerSP := 2, [7].Override := 1, [7].Disable := 1, [7].HI := 100.0, [7].HIHI := 100.0, [7].HITimer.PRE := 5000, [7].HITimerSP := 5, [7].HIHITimer.PRE := 5000, [7].HIHITImerSP := 5, [8].Override := 1, [8].Disable := 1, [8].HITimer.ACC := 100, [8].HITimer.EN := 1, [8].HITimer.DN := 1, [8].HIHITimer.ACC := 100, [8].HIHITimer.EN := 1, [8].HIHITimer.DN := 1, [9].Override := 1, [9].Disable := 1, [9].HITimer.PRE := 60000, [9].HIHITimer.PRE := 60000, [10].Override := 1, [10].Disable := 1, [11].Override := 1, [11].Disable := 1, [11].HITimer.PRE := 60000, [11].HIHITimer.PRE := 20000, [12].Override := 1, [12].Disable := 1, [13].Override := 1, [13].Disable := 1, [14].Override := 1, [14].Disable := 1, [15].Override := 1, [15].Disable := 1, [16].Override := 1, [16].Disable := 1, [17].Override := 1, [17].Disable := 1, [18].Override := 1, [18].Disable := 1, [19].Override := 1, [19].Disable := 1);   // Control Loop Deviation Alarm Array
        [7]   // Mixing Closed Loop Conductivity Deviation Alarm
        [2]   // FI002 Secondary Feed Pump Flow Deviation
        [3]   // Position PCV032 Deviation Alarm
        [1]   // FI001 Primary Feed Pump Flow Deviation
        [6]   // Mixing Closed Loop TotalFlow Deviation Alarm
   AlarmDeviation_Storage : AlarmDeviation[6,20] := ([0,0].Override := 1, [0,0].Disable := 1, [0,0].HIAlarmONS := 1, [0,0].HIHIAlarmONS := 1, [0,0].HI := 40.0, [0,0].HIHI := 53.0, [0,0].LOLOLim := 31.333328, [0,0].LOLim := 39.999992, [0,0].HILim := 93.33332, [0,0].HIHILim := 101.999985, [0,0].HITimer.PRE := 30000, [0,0].HIHITimer.PRE := 30000, [0,1].Override := 1, [0,1].Disable := 1, [0,1].HI := 100.0, [0,1].HIHI := 100.0, [0,1].HITimer.PRE := 5000, [0,1].HITimerSP := 5, [0,1].HIHITimer.PRE := 5000, [0,1].HIHITImerSP := 5, [0,1].EnableCfg := 1, [0,2].Override := 1, [0,2].Disable := 1, [0,2].HI := 100.0, [0,2].HIHI := 100.0, [0,2].HITimer.PRE := 5000, [0,2].HITimerSP := 5, [0,2].HIHITimer.PRE := 5000, [0,2].HIHITImerSP := 5, [0,2].EnableCfg := 1, [0,3].Override := 1, [0,3].Disable := 1, [0,3].HI := 100.0, [0,3].HIHI := 100.0, [0,3].HITimer.PRE := 5000, [0,3].HITimerSP := 5, [0,3].HIHITimer.PRE := 5000, [0,3].HIHITImerSP := 5, [0,3].EnableCfg := 1, [0,4].Override := 1, [0,4].Disable := 1, [0,4].HITimer.PRE := 1000, [0,4].HITimer.ACC := 1086, [0,4].HITimer.EN := 1, [0,4].HITimer.DN := 1, [0,4].HIHITimer.PRE := 1000, [0,4].HIHITimer.ACC := 1086, [0,4].HIHITimer.EN := 1, [0,4].HIHITimer.DN := 1, [0,5].Override := 1, [0,5].Disable := 1, [0,5].HITimer.PRE := 2000, [0,5].HIHITimer.PRE := 2000, [0,6].Override := 1, [0,6].Disable := 1, [0,6].HI := 100.0, [0,6].HIHI := 100.0, [0,6].HILim := 40.0, [0,6].HIHILim := 40.0, [0,6].HITimer.PRE := 5000,
        [0,6].HITimerSP := 5, [0,6].HIHITimer.PRE := 5000, [0,6].HIHITImerSP := 5, [0,6].EnableCfg := 1, [0,7].Override := 1, [0,7].Disable := 1, [0,7].HI := 100.0, [0,7].HIHI := 100.0, [0,7].HITimer.PRE := 5000, [0,7].HITimerSP := 5, [0,7].HIHITimer.PRE := 5000, [0,7].HIHITImerSP := 5, [0,7].EnableCfg := 1, [0,8].Override := 1, [0,8].Disable := 1, [0,8].HITimer.ACC := 100, [0,8].HITimer.EN := 1, [0,8].HITimer.DN := 1, [0,8].HIHITimer.ACC := 100, [0,8].HIHITimer.EN := 1, [0,8].HIHITimer.DN := 1, [0,9].Override := 1, [0,9].Disable := 1, [0,9].HITimer.PRE := 60000, [0,9].HIHITimer.PRE := 60000, [0,10].Override := 1, [0,10].Disable := 1, [0,11].Override := 1, [0,11].Disable := 1, [0,11].HITimer.PRE := 60000, [0,11].HIHITimer.PRE := 20000, [0,12].Override := 1, [0,12].Disable := 1, [0,13].Override := 1, [0,13].Disable := 1, [0,14].Override := 1, [0,14].Disable := 1, [0,15].Override := 1, [0,15].Disable := 1, [0,16].Override := 1, [0,16].Disable := 1, [0,17].Override := 1, [0,17].Disable := 1, [0,18].Override := 1, [0,18].Disable := 1, [0,19].Override := 1, [0,19].Disable := 1, [1,0].Override := 1, [1,0].Disable := 1, [1,0].HIAlarmONS := 1, [1,0].HIHIAlarmONS := 1, [1,0].HI := 40.0, [1,0].HIHI := 53.0, [1,0].LOLOLim := 31.333328, [1,0].LOLim := 39.999992, [1,0].HILim := 93.33332, [1,0].HIHILim := 101.999985, [1,0].HITimer.PRE := 30000, [1,0].HIHITimer.PRE := 30000, [1,1].Override := 1,
        [1,1].Disable := 1, [1,1].HI := 100.0, [1,1].HIHI := 100.0, [1,1].HITimer.PRE := 2000, [1,1].HITimerSP := 2, [1,1].HIHITimer.PRE := 2000, [1,1].HIHITImerSP := 2, [1,1].EnableCfg := 1, [1,2].Override := 1, [1,2].Disable := 1, [1,2].HI := 100.0, [1,2].HIHI := 100.0, [1,2].HITimer.PRE := 2000, [1,2].HITimerSP := 2, [1,2].HIHITimer.PRE := 2000, [1,2].HIHITImerSP := 2, [1,2].EnableCfg := 1, [1,3].Override := 1, [1,3].Disable := 1, [1,3].HI := 100.0, [1,3].HIHI := 100.0, [1,3].HITimer.PRE := 5000, [1,3].HITimerSP := 5, [1,3].HIHITimer.PRE := 5000, [1,3].HIHITImerSP := 5, [1,3].EnableCfg := 1, [1,4].Override := 1, [1,4].Disable := 1, [1,4].HI := 100.0, [1,4].HIHI := 100.0, [1,4].HITimer.PRE := 2000, [1,4].HITimerSP := 2, [1,4].HIHITimer.PRE := 2000, [1,4].HIHITImerSP := 2, [1,5].Override := 1, [1,5].Disable := 1, [1,5].EnableCfg := 1, [1,6].Override := 1, [1,6].Disable := 1, [1,6].HI := 100.0, [1,6].HIHI := 100.0, [1,6].HITimer.PRE := 2000, [1,6].HITimerSP := 2, [1,6].HIHITimer.PRE := 2000, [1,6].HIHITImerSP := 2, [1,7].Override := 1, [1,7].Disable := 1, [1,7].HI := 100.0, [1,7].HIHI := 100.0, [1,7].HITimer.PRE := 5000, [1,7].HITimerSP := 5, [1,7].HIHITimer.PRE := 5000, [1,7].HIHITImerSP := 5, [1,8].Override := 1, [1,8].Disable := 1, [1,8].HITimer.ACC := 100, [1,8].HITimer.EN := 1, [1,8].HITimer.DN := 1, [1,8].HIHITimer.ACC := 100, [1,8].HIHITimer.EN := 1,
        [1,8].HIHITimer.DN := 1, [1,9].Override := 1, [1,9].Disable := 1, [1,9].HITimer.PRE := 60000, [1,9].HIHITimer.PRE := 60000, [1,10].Override := 1, [1,10].Disable := 1, [1,11].Override := 1, [1,11].Disable := 1, [1,11].HITimer.PRE := 60000, [1,11].HIHITimer.PRE := 20000, [1,12].Override := 1, [1,12].Disable := 1, [1,13].Override := 1, [1,13].Disable := 1, [1,14].Override := 1, [1,14].Disable := 1, [1,15].Override := 1, [1,15].Disable := 1, [1,16].Override := 1, [1,16].Disable := 1, [1,17].Override := 1, [1,17].Disable := 1, [1,18].Override := 1, [1,18].Disable := 1, [1,19].Override := 1, [1,19].Disable := 1, [2,0].Override := 1, [2,0].Disable := 1, [2,0].HIAlarmONS := 1, [2,0].HIHIAlarmONS := 1, [2,0].HI := 40.0, [2,0].HIHI := 53.0, [2,0].LOLOLim := 31.33333, [2,0].LOLim := 39.99999, [2,0].HILim := 93.33332, [2,0].HIHILim := 102.0, [2,0].HITimer.PRE := 30000, [2,0].HIHITimer.PRE := 30000, [2,1].Disable := 1, [2,1].HI := 100.0, [2,1].HIHI := 100.0, [2,1].HITimer.PRE := 2000, [2,1].HITimerSP := 2, [2,1].HIHITimer.PRE := 2000, [2,1].HIHITImerSP := 2, [2,1].EnableCfg := 1, [2,2].Disable := 1, [2,2].HI := 100.0, [2,2].HIHI := 100.0, [2,2].HITimer.PRE := 2000, [2,2].HITimerSP := 2, [2,2].HIHITimer.PRE := 2000, [2,2].HIHITImerSP := 2, [2,2].EnableCfg := 1, [2,3].Override := 1, [2,3].Disable := 1, [2,3].HI := 100.0, [2,3].HIHI := 100.0, [2,3].LOLOLim := -100.0,
        [2,3].LOLim := -100.0, [2,3].HILim := 100.0, [2,3].HIHILim := 100.0, [2,3].HITimer.PRE := 5000, [2,3].HITimerSP := 5, [2,3].HIHITimer.PRE := 5000, [2,3].HIHITImerSP := 5, [2,4].HI := 100.0, [2,4].HIHI := 100.0, [2,4].HITimer.PRE := 2000, [2,4].HITimerSP := 2, [2,4].HIHITimer.PRE := 2000, [2,4].HIHITImerSP := 2, [2,4].EnableCfg := 1, [2,5].Override := 1, [2,5].Disable := 1, [2,5].HITimer.PRE := 2000, [2,5].HIHITimer.PRE := 2000, [2,6].HI := 100.0, [2,6].HIHI := 100.0, [2,6].HITimer.PRE := 2000, [2,6].HITimerSP := 2, [2,6].HIHITimer.PRE := 2000, [2,6].HIHITImerSP := 2, [2,6].EnableCfg := 1, [2,7].Disable := 1, [2,7].HI := 100.0, [2,7].HIHI := 100.0, [2,7].HITimer.PRE := 5000, [2,7].HITimerSP := 5, [2,7].HIHITimer.PRE := 5000, [2,7].HIHITImerSP := 5, [2,7].EnableCfg := 1, [2,8].Override := 1, [2,8].Disable := 1, [2,8].HITimer.ACC := 100, [2,8].HITimer.EN := 1, [2,8].HITimer.DN := 1, [2,8].HIHITimer.ACC := 100, [2,8].HIHITimer.EN := 1, [2,8].HIHITimer.DN := 1, [2,9].Override := 1, [2,9].Disable := 1, [2,9].HITimer.PRE := 60000, [2,9].HIHITimer.PRE := 60000, [2,10].Override := 1, [2,10].Disable := 1, [2,11].Override := 1, [2,11].Disable := 1, [2,11].HITimer.PRE := 60000, [2,11].HIHITimer.PRE := 20000, [2,12].Override := 1, [2,12].Disable := 1, [2,13].Override := 1, [2,13].Disable := 1, [2,14].Override := 1, [2,14].Disable := 1, [2,15].Override := 1, [2,15].Disable := 1, [2,16].Override := 1,
        [2,16].Disable := 1, [2,17].Override := 1, [2,17].Disable := 1, [2,18].Override := 1, [2,18].Disable := 1, [2,19].Override := 1, [2,19].Disable := 1, [3,0].Override := 1, [3,0].Disable := 1, [3,1].Disable := 1, [3,1].EnableCfg := 1, [3,2].Disable := 1, [3,2].EnableCfg := 1, [3,3].HIAlarm := 1, [3,3].HIHIAlarm := 1, [3,3].HIAlarmONS := 1, [3,3].HIHIAlarmONS := 1, [3,3].HITimer.EN := 1, [3,3].HITimer.DN := 1, [3,3].HIHITimer.EN := 1, [3,3].HIHITimer.DN := 1, [3,3].EnableCfg := 1, [3,4].Override := 1, [3,4].Disable := 1, [3,5].Override := 1, [3,5].Disable := 1, [3,6].Disable := 1, [3,6].EnableCfg := 1, [3,7].Disable := 1, [3,7].EnableCfg := 1, [3,8].Override := 1, [3,8].Disable := 1, [3,9].Override := 1, [3,9].Disable := 1, [3,10].Override := 1, [3,10].Disable := 1, [3,11].Override := 1, [3,11].Disable := 1, [3,12].Override := 1, [3,12].Disable := 1, [3,13].Override := 1, [3,13].Disable := 1, [3,14].Override := 1, [3,14].Disable := 1, [3,15].Override := 1, [3,15].Disable := 1, [3,16].Override := 1, [3,16].Disable := 1, [3,17].Override := 1, [3,17].Disable := 1, [3,18].Override := 1, [3,18].Disable := 1, [3,19].Override := 1, [3,19].Disable := 1, [4,0].Override := 1, [4,0].Disable := 1, [4,0].HIAlarmONS := 1, [4,0].HIHIAlarmONS := 1, [4,0].HI := 40.0, [4,0].HIHI := 53.0,
        [4,0].LOLOLim := 31.333328, [4,0].LOLim := 39.999992, [4,0].HILim := 93.33332, [4,0].HIHILim := 101.999985, [4,0].HITimer.PRE := 30000, [4,0].HIHITimer.PRE := 30000, [4,1].Override := 1, [4,1].Disable := 1, [4,1].HI := 100.0, [4,1].HIHI := 100.0, [4,1].HITimer.PRE := 5000, [4,1].HITimerSP := 5, [4,1].HIHITimer.PRE := 5000, [4,1].HIHITImerSP := 5, [4,1].EnableCfg := 1, [4,2].Override := 1, [4,2].Disable := 1, [4,2].HI := 100.0, [4,2].HIHI := 100.0, [4,2].HITimer.PRE := 5000, [4,2].HITimerSP := 5, [4,2].HIHITimer.PRE := 5000, [4,2].HIHITImerSP := 5, [4,2].EnableCfg := 1, [4,3].Override := 1, [4,3].Disable := 1, [4,3].HI := 20.0, [4,3].HIHI := 30.0, [4,3].LOLOLim := -30.0, [4,3].LOLim := -20.0, [4,3].HILim := 20.0, [4,3].HIHILim := 30.0, [4,3].HITimer.PRE := 5000, [4,3].HITimerSP := 5, [4,3].HIHITimer.PRE := 5000, [4,3].HIHITImerSP := 5, [4,3].EnableCfg := 1, [4,4].Override := 1, [4,4].Disable := 1, [4,4].HITimer.PRE := 1000, [4,4].HITimer.ACC := 1086, [4,4].HITimer.EN := 1, [4,4].HITimer.DN := 1, [4,4].HIHITimer.PRE := 1000, [4,4].HIHITimer.ACC := 1086, [4,4].HIHITimer.EN := 1, [4,4].HIHITimer.DN := 1, [4,5].Override := 1, [4,5].Disable := 1, [4,5].HITimer.PRE := 2000, [4,5].HIHITimer.PRE := 2000, [4,6].Override := 1, [4,6].Disable := 1, [4,6].HI := 100.0, [4,6].HIHI := 100.0, [4,6].LOLOLim := 5.0, [4,6].LOLim := 5.0, [4,6].HILim := 15.0, [4,6].HIHILim := 15.0, [4,6].HITimer.PRE := 5000,
        [4,6].HITimerSP := 5, [4,6].HIHITimer.PRE := 5000, [4,6].HIHITImerSP := 5, [4,6].EnableCfg := 1, [4,7].Override := 1, [4,7].Disable := 1, [4,7].HI := 100.0, [4,7].HIHI := 100.0, [4,7].HITimer.PRE := 5000, [4,7].HITimerSP := 5, [4,7].HIHITimer.PRE := 5000, [4,7].HIHITImerSP := 5, [4,7].EnableCfg := 1, [4,8].Override := 1, [4,8].Disable := 1, [4,8].HITimer.ACC := 100, [4,8].HITimer.EN := 1, [4,8].HITimer.DN := 1, [4,8].HIHITimer.ACC := 100, [4,8].HIHITimer.EN := 1, [4,8].HIHITimer.DN := 1, [4,9].Override := 1, [4,9].Disable := 1, [4,9].HITimer.PRE := 60000, [4,9].HIHITimer.PRE := 60000, [4,10].Override := 1, [4,10].Disable := 1, [4,11].Override := 1, [4,11].Disable := 1, [4,11].HITimer.PRE := 60000, [4,11].HIHITimer.PRE := 20000, [4,12].Override := 1, [4,12].Disable := 1, [4,13].Override := 1, [4,13].Disable := 1, [4,14].Override := 1, [4,14].Disable := 1, [4,15].Override := 1, [4,15].Disable := 1, [4,16].Override := 1, [4,16].Disable := 1, [4,17].Override := 1, [4,17].Disable := 1, [4,18].Override := 1, [4,18].Disable := 1, [4,19].Override := 1, [4,19].Disable := 1, [5,0].Override := 1, [5,0].Disable := 1, [5,0].HIAlarmONS := 1, [5,0].HIHIAlarmONS := 1, [5,0].HI := 40.0, [5,0].HIHI := 53.0, [5,0].LOLOLim := 31.333328, [5,0].LOLim := 39.999992, [5,0].HILim := 93.33332, [5,0].HIHILim := 101.999985, [5,0].HITimer.PRE := 30000, [5,0].HIHITimer.PRE := 30000, [5,1].Override := 1,
        [5,1].Disable := 1, [5,1].HI := 100.0, [5,1].HIHI := 100.0, [5,1].HITimer.PRE := 5000, [5,1].HITimerSP := 5, [5,1].HIHITimer.PRE := 5000, [5,1].HIHITImerSP := 5, [5,1].EnableCfg := 1, [5,2].Override := 1, [5,2].Disable := 1, [5,2].HI := 100.0, [5,2].HIHI := 100.0, [5,2].HITimer.PRE := 5000, [5,2].HITimerSP := 5, [5,2].HIHITimer.PRE := 5000, [5,2].HIHITImerSP := 5, [5,2].EnableCfg := 1, [5,3].Override := 1, [5,3].Disable := 1, [5,3].HI := 100.0, [5,3].HIHI := 100.0, [5,3].HITimer.PRE := 5000, [5,3].HITimerSP := 5, [5,3].HIHITimer.PRE := 5000, [5,3].HIHITImerSP := 5, [5,3].EnableCfg := 1, [5,4].Override := 1, [5,4].Disable := 1, [5,4].HITimer.PRE := 1000, [5,4].HITimer.ACC := 1086, [5,4].HITimer.EN := 1, [5,4].HITimer.DN := 1, [5,4].HIHITimer.PRE := 1000, [5,4].HIHITimer.ACC := 1086, [5,4].HIHITimer.EN := 1, [5,4].HIHITimer.DN := 1, [5,5].Override := 1, [5,5].Disable := 1, [5,5].HITimer.PRE := 2000, [5,5].HIHITimer.PRE := 2000, [5,6].Override := 1, [5,6].Disable := 1, [5,6].HI := 100.0, [5,6].HIHI := 100.0, [5,6].LOLOLim := 5.0, [5,6].LOLim := 5.0, [5,6].HILim := 15.0, [5,6].HIHILim := 15.0, [5,6].HITimer.PRE := 5000, [5,6].HITimerSP := 5, [5,6].HIHITimer.PRE := 5000, [5,6].HIHITImerSP := 5, [5,6].EnableCfg := 1, [5,7].Override := 1, [5,7].Disable := 1, [5,7].HI := 100.0, [5,7].HIHI := 100.0, [5,7].HITimer.PRE := 5000, [5,7].HITimerSP := 5, [5,7].HIHITimer.PRE := 5000,
        [5,7].HIHITImerSP := 5, [5,7].EnableCfg := 1, [5,8].Override := 1, [5,8].Disable := 1, [5,8].HITimer.ACC := 100, [5,8].HITimer.EN := 1, [5,8].HITimer.DN := 1, [5,8].HIHITimer.ACC := 100, [5,8].HIHITimer.EN := 1, [5,8].HIHITimer.DN := 1, [5,9].Override := 1, [5,9].Disable := 1, [5,9].HITimer.PRE := 60000, [5,9].HIHITimer.PRE := 60000, [5,10].Override := 1, [5,10].Disable := 1, [5,11].Override := 1, [5,11].Disable := 1, [5,11].HITimer.PRE := 60000, [5,11].HIHITimer.PRE := 20000, [5,12].Override := 1, [5,12].Disable := 1, [5,13].Override := 1, [5,13].Disable := 1, [5,14].Override := 1, [5,14].Disable := 1, [5,15].Override := 1, [5,15].Disable := 1, [5,16].Override := 1, [5,16].Disable := 1, [5,17].Override := 1, [5,17].Disable := 1, [5,18].Override := 1, [5,18].Disable := 1, [5,19].Override := 1, [5,19].Disable := 1);
   AnalogOutput : AnalogOutput[25] := ([0].Tag := 'PCV001_AO', [0].RawValue := 47, [0].RawMax := 2047, [0].ScaledValue := 2.2879825, [0].ScaledMax := 100.0, [0].EnableCfg := 1, [1].Tag := 'PCV101_AO', [1].RawValue := 1768, [1].RawMax := 2047, [1].ScaledValue := 86.3938, [1].ScaledMax := 100.0, [1].EnableCfg := 1, [2].Tag := 'SIC001_AO', [2].RawMax := 27648, [2].ScaledMax := 100.0, [2].EnableCfg := 1, [3].Tag := 'SIC002_AO', [3].RawMax := 27648, [3].ScaledMax := 100.0, [3].EnableCfg := 1, [4].Tag := 'SIC003_AO', [4].RawMax := 2047, [4].ScaledMax := 100.0, [4].EnableCfg := 1, [5].Tag := 'SPARE', [5].RawMax := 27648, [5].ScaledMax := 100.0, [6].Tag := 'SPARE', [6].RawValue := -6912, [6].RawMax := 27648, [6].ScaledValue := -25.0, [6].ScaledMax := 100.0, [7].Tag := 'SPARE', [7].RawMax := 27648, [7].ScaledMax := 100.0, [8].Tag := 'AO#1', [8].RawMax := 2047, [8].ScaledMax := 100.0, [9].Tag := 'AO#2', [9].RawMax := 2047, [9].ScaledMax := 100.0, [10].Tag := 'AO#3', [10].RawMax := 2047, [10].ScaledMax := 100.0, [11].Tag := 'AO#4', [11].RawMax := 2047, [11].ScaledMax := 100.0);   // Analog Output Array
        [0]   // Retentate Pressure Control Valve Setpoint
        [1]   // FiltratePressure Control Valve Setpoint
        [4]   // Mixer Speed Setpoint
        [3]   // Transfer Pump Speed Setpoint
        [2]   // Feed Pump Speed Setpoint
   AnalogOutput_Storage : AnalogOutput[6,25] := ([0,0].Tag := 'SIC001', [0,0].RawMax := 27648, [0,0].ScaledMax := 100.0, [0,0].EnableCfg := 1, [0,1].Tag := 'SIC002', [0,1].RawMax := 27648, [0,1].ScaledMax := 100.0, [0,1].EnableCfg := 1, [0,2].Tag := 'PCV010', [0,2].RawMax := 2047, [0,2].ScaledMax := 100.0, [0,2].EnableCfg := 1, [0,3].Tag := 'PCV011', [0,3].RawMax := 27648, [0,3].ScaledMax := 100.0, [0,4].Tag := 'PCV012', [0,4].RawMax := 27648, [0,4].ScaledMax := 100.0, [0,5].Tag := 'SPARE', [0,5].RawMax := 27648, [0,5].ScaledMax := 100.0, [0,6].Tag := 'SPARE', [0,6].RawValue := -6912, [0,6].RawMax := 27648, [0,6].ScaledValue := -25.0, [0,6].ScaledMax := 100.0, [0,7].Tag := 'SPARE', [0,7].RawMax := 27648, [0,7].ScaledMax := 100.0, [0,8].Tag := 'AO#1', [0,8].RawMax := 2047, [0,8].ScaledMax := 100.0, [0,8].EnableCfg := 1, [0,9].Tag := 'AO#2', [0,9].RawMax := 2047, [0,9].ScaledMax := 100.0, [0,9].EnableCfg := 1, [0,10].Tag := 'AO#3', [0,10].RawMax := 2047, [0,10].ScaledMax := 100.0, [0,10].EnableCfg := 1, [0,11].Tag := 'AO#4', [0,11].RawMax := 2047, [0,11].ScaledMax := 100.0, [0,11].EnableCfg := 1, [1,0].Tag := 'PCV001_AO', [1,0].RawMax := 2047, [1,0].ScaledMax := 100.0, [1,0].EnableCfg := 1, [1,1].Tag := 'PCV101_AO', [1,1].RawMax := 2047, [1,1].ScaledMax := 100.0, [1,1].EnableCfg := 1, [1,2].Tag := 'SIC001_AO', [1,2].RawMax := 27648, [1,2].ScaledMax := 100.0, [1,2].EnableCfg := 1, [1,3].Tag := 'SIC002_AO', [1,3].RawMax := 27648, [1,3].ScaledMax := 100.0,
        [1,3].EnableCfg := 1, [1,4].Tag := 'SIC003_AO', [1,4].RawMax := 2047, [1,4].ScaledMax := 100.0, [1,4].EnableCfg := 1, [1,5].Tag := 'SPARE', [1,5].RawMax := 27648, [1,5].ScaledMax := 100.0, [1,6].Tag := 'SPARE', [1,6].RawValue := -6912, [1,6].RawMax := 27648, [1,6].ScaledValue := -25.0, [1,6].ScaledMax := 100.0, [1,7].Tag := 'SPARE', [1,7].RawMax := 27648, [1,7].ScaledMax := 100.0, [1,8].Tag := 'AO#1', [1,8].RawMax := 2047, [1,8].ScaledMax := 100.0, [1,9].Tag := 'AO#2', [1,9].RawMax := 2047, [1,9].ScaledMax := 100.0, [1,10].Tag := 'AO#3', [1,10].RawMax := 2047, [1,10].ScaledMax := 100.0, [1,11].Tag := 'AO#4', [1,11].RawMax := 2047, [1,11].ScaledMax := 100.0, [2,0].Tag := 'PCV001_AO', [2,0].RawMax := 2047, [2,0].ScaledMax := 100.0, [2,0].EnableCfg := 1, [2,1].Tag := 'PCV101_AO', [2,1].RawMax := 2047, [2,1].ScaledMax := 100.0, [2,1].EnableCfg := 1, [2,2].Tag := 'SIC001_AO', [2,2].RawMax := 27648, [2,2].ScaledMax := 100.0, [2,2].EnableCfg := 1, [2,3].Tag := 'SIC002_AO', [2,3].RawMax := 27648, [2,3].ScaledMax := 100.0, [2,3].EnableCfg := 1, [2,4].Tag := 'SIC003_AO', [2,4].RawMax := 2047, [2,4].ScaledMax := 100.0, [2,4].EnableCfg := 1, [2,5].Tag := 'SPARE', [2,5].RawMax := 27648, [2,5].ScaledMax := 100.0, [2,6].Tag := 'SPARE', [2,6].RawValue := -6912, [2,6].RawMax := 27648, [2,6].ScaledValue := -25.0, [2,6].ScaledMax := 100.0, [2,7].Tag := 'SPARE', [2,7].RawMax := 27648, [2,7].ScaledMax := 100.0, [2,8].Tag := 'AO#1',
        [2,8].RawMax := 2047, [2,8].ScaledMax := 100.0, [2,9].Tag := 'AO#2', [2,9].RawMax := 2047, [2,9].ScaledMax := 100.0, [2,10].Tag := 'AO#3', [2,10].RawMax := 2047, [2,10].ScaledMax := 100.0, [2,11].Tag := 'AO#4', [2,11].RawMax := 2047, [2,11].ScaledMax := 100.0, [3,0].RawMax := 27648, [3,0].ScaledMax := 100.0, [3,0].EnableCfg := 1, [3,1].RawMax := 27648, [3,1].ScaledMax := 100.0, [3,1].EnableCfg := 1, [3,2].RawMax := 2047, [3,2].ScaledMax := 100.0, [3,2].EnableCfg := 1, [3,3].RawMax := 27648, [3,3].ScaledMax := 100.0, [3,4].RawMax := 27648, [3,4].ScaledMax := 100.0, [3,5].RawMax := 27648, [3,5].ScaledMax := 100.0, [3,6].RawMax := 27648, [3,6].ScaledMax := 100.0, [3,7].RawMax := 27648, [3,7].ScaledMax := 100.0, [3,8].RawMax := 2047, [3,8].ScaledMax := 100.0, [3,8].EnableCfg := 1, [3,9].RawMax := 2047, [3,9].ScaledMax := 100.0, [3,9].EnableCfg := 1, [3,10].RawMax := 2047, [3,10].ScaledMax := 100.0, [3,10].EnableCfg := 1, [3,11].RawMax := 2047, [3,11].ScaledMax := 100.0, [3,11].EnableCfg := 1, [4,0].Tag := 'SIC001', [4,0].RawMax := 27648, [4,0].ScaledMax := 100.0, [4,0].EnableCfg := 1, [4,1].Tag := 'SIC002', [4,1].RawMax := 27648, [4,1].ScaledMax := 100.0, [4,1].EnableCfg := 1, [4,2].Tag := 'PCV010', [4,2].RawMax := 2047, [4,2].ScaledMax := 100.0, [4,2].EnableCfg := 1, [4,3].Tag := 'PCV011', [4,3].RawMax := 27648, [4,3].ScaledMax := 100.0, [4,4].Tag := 'PCV012', [4,4].RawMax := 27648, [4,4].ScaledMax := 100.0,
        [4,5].Tag := 'SPARE', [4,5].RawMax := 27648, [4,5].ScaledMax := 100.0, [4,6].Tag := 'SPARE', [4,6].RawValue := -6912, [4,6].RawMax := 27648, [4,6].ScaledValue := -25.0, [4,6].ScaledMax := 100.0, [4,7].Tag := 'SPARE', [4,7].RawMax := 27648, [4,7].ScaledMax := 100.0, [4,8].Tag := 'AO#1', [4,8].RawMax := 2047, [4,8].ScaledMax := 100.0, [4,8].EnableCfg := 1, [4,9].Tag := 'AO#2', [4,9].RawMax := 2047, [4,9].ScaledMax := 100.0, [4,9].EnableCfg := 1, [4,10].Tag := 'AO#3', [4,10].RawMax := 2047, [4,10].ScaledMax := 100.0, [4,10].EnableCfg := 1, [4,11].Tag := 'AO#4', [4,11].RawMax := 2047, [4,11].ScaledMax := 100.0, [4,11].EnableCfg := 1, [5,0].Tag := 'SIC001', [5,0].RawMax := 27648, [5,0].ScaledMax := 100.0, [5,0].EnableCfg := 1, [5,1].Tag := 'SIC002', [5,1].RawMax := 27648, [5,1].ScaledMax := 100.0, [5,1].EnableCfg := 1, [5,2].Tag := 'PCV010', [5,2].RawMax := 2047, [5,2].ScaledMax := 100.0, [5,2].EnableCfg := 1, [5,3].Tag := 'PCV011', [5,3].RawMax := 27648, [5,3].ScaledMax := 100.0, [5,4].Tag := 'PCV012', [5,4].RawMax := 27648, [5,4].ScaledMax := 100.0, [5,5].Tag := 'SPARE', [5,5].RawMax := 27648, [5,5].ScaledMax := 100.0, [5,6].Tag := 'SPARE', [5,6].RawValue := -6912, [5,6].RawMax := 27648, [5,6].ScaledValue := -25.0, [5,6].ScaledMax := 100.0, [5,7].Tag := 'SPARE', [5,7].RawMax := 27648, [5,7].ScaledMax := 100.0, [5,8].Tag := 'AO#1', [5,8].RawMax := 2047, [5,8].ScaledMax := 100.0, [5,8].EnableCfg := 1,
        [5,9].Tag := 'AO#2', [5,9].RawMax := 2047, [5,9].ScaledMax := 100.0, [5,9].EnableCfg := 1, [5,10].Tag := 'AO#3', [5,10].RawMax := 2047, [5,10].ScaledMax := 100.0, [5,10].EnableCfg := 1, [5,11].Tag := 'AO#4', [5,11].RawMax := 2047, [5,11].ScaledMax := 100.0, [5,11].EnableCfg := 1);
   AnalogPoint : AnalogInput[50] := ([0].TagName := 'WI101', [0].RawMax := 99999, [0].RawLowLimit := -1000, [0].RawHighLimit := 100999, [0].FilterActual := 1.0, [0].ScaledMax := 9999.9, [0].RangeMax := 1500.0, [0].RangeMaxSave := 1500.0, [0].OverrideCfg := 1, [0].EGU := 'kg', [1].TagName := 'WI102', [1].OutofRange := 1, [1].Address := 1, [1].RawMin := 6553, [1].RawMax := 32767, [1].RawValue := 1, [1].RawLowLimit := 6225, [1].RawHighLimit := 33095, [1].FilterActual := 1.0, [1].ScaledMax := 1500.0, [1].CurrentValue := -374.9619, [1].RangeMax := 1500.0, [1].RangeMaxSave := 1500.0, [1].EnableCfg := 1, [1].OverrideCfg := 1, [1].EGU := 'kg', [2].TagName := 'FI101', [2].Address := 2, [2].RawMin := 6553, [2].RawMax := 32767, [2].RawLowLimit := 6225, [2].RawHighLimit := 33095, [2].FilterActual := 1.0, [2].ScaledMax := 20.0, [2].RangeMax := 25.0, [2].RangeMaxSave := 25.0, [2].EnableCfg := 1, [2].OverrideCfg := 1, [2].EGU := 'Lpm', [3].TagName := 'PCV001', [3].Address := 3, [3].RawMin := 6553, [3].RawMax := 32767, [3].RawValue := 23484, [3].RawLowLimit := 6225, [3].RawHighLimit := 33095, [3].FilteredRaw := 23484, [3].FilterActual := 1.0, [3].ScaledMax := 100.0, [3].CurrentValue := -0.03292181, [3].RangeMax := 100.0, [3].RangeMaxSave := 100.0, [3].EnableCfg := 1, [3].EGU := '%Clo', [4].TagName := 'PCV101', [4].Address := 4, [4].RawMin := 6553, [4].RawMax := 32767, [4].RawValue := 23322, [4].RawLowLimit := 6225,
        [4].RawHighLimit := 33095, [4].FilteredRaw := 23322, [4].FilterActual := 1.0, [4].ScaledMax := 100.0, [4].CurrentValue := 99.47403, [4].RangeMax := 100.0, [4].RangeMaxSave := 100.0, [4].EnableCfg := 1, [4].EGU := '%Opn', [5].TagName := 'PI001', [5].Address := 5, [5].RawMin := 6553, [5].RawMax := 32767, [5].RawValue := 6577, [5].RawLowLimit := 6225, [5].RawHighLimit := 33095, [5].FilteredRaw := 6577, [5].FilterActual := 1.0, [5].ScaledMax := 87.0, [5].CurrentValue := 0.0796521, [5].RangeMax := 87.0, [5].RangeMaxSave := 87.0, [5].RealCfg := 1, [5].EnableCfg := 1, [5].OverrideCfg := 1, [5].EGU := 'psi', [6].TagName := 'PI002', [6].Address := 6, [6].RawMin := 6553, [6].RawMax := 32767, [6].RawValue := 6476, [6].RawLowLimit := 6225, [6].RawHighLimit := 33095, [6].FilterUser := 50, [6].FilteredRaw := 6484, [6].FilterActual := 0.5, [6].ScaledMax := 87.0, [6].CurrentValue := -0.22899978, [6].RangeMax := 87.0, [6].RangeMaxSave := 87.0, [6].RealCfg := 1, [6].EnableCfg := 1, [6].OverrideCfg := 1, [6].EGU := 'psi', [7].TagName := 'PI101', [7].Address := 7, [7].RawMin := 6553, [7].RawMax := 32767, [7].RawValue := 6504, [7].RawLowLimit := 6225, [7].RawHighLimit := 33095, [7].FilteredRaw := 6504, [7].FilterActual := 1.0, [7].ScaledMax := 87.0, [7].CurrentValue := -0.16262303, [7].RangeMax := 87.0, [7].RangeMaxSave := 87.0, [7].RealCfg := 1, [7].EnableCfg := 1, [7].OverrideCfg := 1,
        [7].EGU := 'psi', [8].TagName := 'PI401', [8].Address := 8, [8].RawMin := 6553, [8].RawMax := 32767, [8].RawValue := 6641, [8].RawLowLimit := 6225, [8].RawHighLimit := 33095, [8].FilteredRaw := 6641, [8].FilterActual := 1.0, [8].ScaledMax := 87.0, [8].CurrentValue := 0.2920577, [8].RangeMax := 87.0, [8].RangeMaxSave := 87.0, [8].RealCfg := 1, [8].EnableCfg := 1, [8].OverrideCfg := 1, [8].EGU := 'psi', [9].TagName := 'AI104', [9].OutofRange := 1, [9].Address := 9, [9].RawMin := 6553, [9].RawMax := 32767, [9].RawLowLimit := 6225, [9].RawHighLimit := 33095, [9].FilterActual := 1.0, [9].ScaledMax := 14.0, [9].CurrentValue := -1.4998856, [9].RangeMax := 14.0, [9].RangeMaxSave := 14.0, [9].RealCfg := 1, [9].OverrideCfg := 1, [9].EGU := 'pH', [10].TagName := 'AI101', [10].Address := 10, [10].RawMin := 6553, [10].RawMax := 32767, [10].RawValue := 6559, [10].RawLowLimit := 6225, [10].RawHighLimit := 33095, [10].FilteredRaw := 6559, [10].FilterActual := 1.0, [10].ScaledMax := 200.0, [10].CurrentValue := 0.045777068, [10].RangeMax := 200.0, [10].RangeMaxSave := 200.0, [10].RealCfg := 1, [10].EnableCfg := 1, [10].OverrideCfg := 1, [10].EGU := 'mS/cm', [11].TagName := 'AI102', [11].Address := 11, [11].RawMin := 6553, [11].RawMax := 32767, [11].RawValue := 7802, [11].RawLowLimit := 6225, [11].RawHighLimit := 33095, [11].FilteredRaw := 7802, [11].FilterActual := 1.0, [11].ScaledMax := 2.0,
        [11].CurrentValue := 0.09529259, [11].RangeMax := 2.0, [11].RangeMaxSave := 2.0, [11].RealCfg := 1, [11].EnableCfg := 1, [11].OverrideCfg := 1, [11].EGU := 'AU', [12].TagName := 'AI103', [12].Address := 12, [12].RawMin := 6553, [12].RawMax := 32767, [12].RawValue := 6959, [12].RawLowLimit := 6225, [12].RawHighLimit := 33095, [12].FilteredRaw := 6959, [12].FilterActual := 1.0, [12].ScaledMax := 2.0, [12].CurrentValue := 0.030975815, [12].RangeMax := 2.0, [12].RangeMaxSave := 2.0, [12].RealCfg := 1, [12].EnableCfg := 1, [12].OverrideCfg := 1, [12].EGU := 'AU', [13].TagName := 'TI001', [13].Address := 13, [13].RawMin := 6553, [13].RawMax := 32767, [13].RawValue := 16343, [13].RawLowLimit := 6225, [13].RawHighLimit := 33095, [13].FilteredRaw := 16343, [13].FilterActual := 1.0, [13].ScaledMax := 55.0, [13].CurrentValue := 20.540552, [13].RangeMax := 55.0, [13].RangeMaxSave := 55.0, [13].RealCfg := 1, [13].EnableCfg := 1, [13].OverrideCfg := 1, [13].EGU := '$B0C', [14].TagName := 'MIX001', [14].Address := 14, [14].RawMax := 16384, [14].RawValue := 45, [14].RawLowLimit := -164, [14].RawHighLimit := 16548, [14].FilteredRaw := 45, [14].FilterActual := 1.0, [14].ScaledMax := 100.0, [14].CurrentValue := 0.2746582, [14].RangeMax := 100.0, [14].RangeMaxSave := 100.0, [14].RealCfg := 1, [14].EnableCfg := 1, [14].EGU := '%', [15].TagName := 'WI001', [15].Address := 15, [15].RawMax := 99999, [15].RawLowLimit := -1000,
        [15].RawHighLimit := 100999, [15].FilterActual := 1.0, [15].ScaledMax := 999.99, [15].EnableCfg := 1, [15].OverrideCfg := 1, [16].CurrentValue := -0.4999322, [17].Address := 17, [17].RawMin := 6553, [17].RawMax := 32767, [17].CurrentValue := -2.499796, [17].RealCfg := 1, [17].OverrideCfg := 1, [18].CurrentValue := -2.499796, [19].CurrentValue := -2.499796, [20].CurrentValue := -24.99661, [21].CurrentValue := -24.99661, [22].TagName := 'SPARE', [23].TagName := 'SPARE', [24].TagName := 'SPARE', [25].TagName := 'SPARE', [26].TagName := 'SPARE', [27].TagName := 'SPARE', [28].TagName := 'AI#1', [28].Address := 28, [28].RawMin := 6553, [28].RawMax := 32767, [28].RawValue := 12544, [28].RawLowLimit := 6225, [28].RawHighLimit := 33095, [28].FilteredRaw := 12544, [28].FilterActual := 1.0, [28].ScaledMax := 100.0, [28].CurrentValue := 22.8542, [28].RangeMax := 100.0, [28].RangeMaxSave := 100.0, [28].RealCfg := 1, [28].OverrideCfg := 1, [29].TagName := 'AI#2', [29].Address := 29, [29].RawMin := 6553, [29].RawMax := 32767, [29].RawValue := 12288, [29].RawLowLimit := 6225, [29].RawHighLimit := 33095, [29].FilteredRaw := 12288, [29].FilterActual := 1.0, [29].ScaledMax := 100.0, [29].CurrentValue := 21.877623, [29].RangeMax := 100.0, [29].RangeMaxSave := 100.0, [29].RealCfg := 1, [29].OverrideCfg := 1, [30].TagName := 'AI#3', [30].Address := 30, [30].RawMin := 6553, [30].RawMax := 32767, [30].RawValue := 12288, [30].RawLowLimit := 6225, [30].RawHighLimit := 33095, [30].FilteredRaw := 12288,
        [30].FilterActual := 1.0, [30].ScaledMax := 100.0, [30].CurrentValue := 21.877623, [30].RangeMax := 100.0, [30].RangeMaxSave := 100.0, [30].RealCfg := 1, [30].OverrideCfg := 1, [31].TagName := 'AI#4', [31].Address := 31, [31].RawMin := 6553, [31].RawMax := 32767, [31].RawValue := 12288, [31].RawLowLimit := 6225, [31].RawHighLimit := 33095, [31].FilteredRaw := 12288, [31].FilterActual := 1.0, [31].ScaledMax := 100.0, [31].CurrentValue := 21.877623, [31].RangeMax := 100.0, [31].RangeMaxSave := 100.0, [31].RealCfg := 1, [31].OverrideCfg := 1, [40].TagName := 'DP', [40].Address := 40, [40].RawMin := 6553, [40].RawMax := 32767, [40].RawLowLimit := 6225, [40].RawHighLimit := 33095, [40].FilterActual := 1.0, [40].ScaledMax := 87.0, [40].CurrentValue := 0.18917373, [40].RangeMax := 87.0, [40].RangeMaxSave := 87.0, [40].EnableCfg := 1, [40].OverrideCfg := 1, [40].EGU := 'psi', [41].TagName := 'TMP', [41].Address := 41, [41].RawMin := 6553, [41].RawMax := 32767, [41].RawLowLimit := 6225, [41].RawHighLimit := 33095, [41].FilterActual := 1.0, [41].ScaledMax := 87.0, [41].CurrentValue := 0.087949194, [41].RangeMax := 87.0, [41].RangeMaxSave := 87.0, [41].EnableCfg := 1, [41].OverrideCfg := 1, [41].EGU := 'psi', [42].TagName := 'FI001', [42].Address := 42, [42].RawMin := 6553, [42].RawMax := 32767, [42].RawLowLimit := 6225, [42].RawHighLimit := 33095, [42].FilterActual := 1.0, [42].ScaledMax := 48.0, [42].RangeMax := 48.0, [42].RangeMaxSave := 48.0,
        [42].EnableCfg := 1, [42].OverrideCfg := 1, [42].EGU := 'Lpm', [43].TagName := 'FI401', [43].Address := 43, [43].RawMin := 6553, [43].RawMax := 32767, [43].RawLowLimit := 6225, [43].RawHighLimit := 33095, [43].FilterActual := 1.0, [43].ScaledMax := 25.0, [43].RangeMax := 25.0, [43].RangeMaxSave := 25.0, [43].EnableCfg := 1, [43].OverrideCfg := 1, [43].EGU := 'Lpm', [44].TagName := 'LI001', [44].Address := 44, [44].RawMin := 6553, [44].RawMax := 32767, [44].RawLowLimit := 6225, [44].RawHighLimit := 33095, [44].FilterActual := 1.0, [44].ScaledMax := 200.0, [44].RangeMax := 200.0, [44].RangeMaxSave := 200.0, [44].EnableCfg := 1, [44].OverrideCfg := 1, [45].TagName := 'NWP', [45].Address := 45, [45].RawMin := 6553, [45].RawMax := 32767, [45].RawLowLimit := 6225, [45].RawHighLimit := 33095, [45].FilterActual := 1.0, [45].ScaledMax := 999.0, [45].RangeMax := 999.0, [45].RangeMaxSave := 999.0, [45].EnableCfg := 1, [45].EGU := 'Lm$B2h/', [46].TagName := 'PERM', [46].Address := 46, [46].RawMin := 6553, [46].RawMax := 32767, [46].RawLowLimit := 6225, [46].RawHighLimit := 33095, [46].FilterActual := 1.0, [46].ScaledMax := 999.0, [46].RangeMax := 999.0, [46].RangeMaxSave := 999.0, [46].EnableCfg := 1, [46].EGU := 'Lm$B2h/');   // Analog Input Array
        [1]   // Customer Filtrate Wheight
        [3]   // Retentate Pressure Control Valve Position
        [4]   // Filtrate Pressure Control Valve Position
        [45]   // Normalized Water Permeability
        [41]   // Trans-Membrane Pressure
        [17]   // Retentate Flow
        [16]   // Filtrate bag Weight
        [6]   // Retentate Pressure
        [11]   // Filtrate UV
        [12]   // Filtrate UV
        [14]   // Mixer Speed
        [2]   // Filtrate Flow
        [5]   // Feed Pressure
        [42]   // Feed Flow
        [9]   // Filtrate pH
        [43]   // Transfer Pump Flow
        [0]   // Filtrate Weight
        [13]   // Feed Bag Temperature
        [15]   // Feed bag Weight
        [8]   // Transfer Pump Pressure
        [44]   // Feed Bag volume
        [10]   // Filtrate Conductivity
        [40]   // Differential Pressure
        [46]   // Membrane Permeability
        [7]   // Filtrate Pressure
   AnalogPoint_Storage : AnalogInput[6,50] := ([0,0].TagName := 'PCV032', [0,0].OutofRange := 1, [0,0].RawMin := 6553, [0,0].RawMax := 32767, [0,0].RawValue := 1, [0,0].RawLowLimit := 6225, [0,0].RawHighLimit := 33095, [0,0].FilteredRaw := 1, [0,0].FilterActual := 1.0, [0,0].ScaledMax := 100.0, [0,0].CurrentValue := -24.994278, [0,0].RangeMax := 100.0, [0,0].RangeMaxSave := 100.0, [0,0].RealCfg := 1, [0,0].EnableCfg := 1, [0,0].OverrideCfg := 1, [0,1].TagName := 'AI201B', [0,1].OutofRange := 1, [0,1].Address := 1, [0,1].RawMin := 5529, [0,1].RawMax := 27648, [0,1].RawLowLimit := 5253, [0,1].RawHighLimit := 27924, [0,1].FilterActual := 1.0, [0,1].ScaledMax := 50.0, [0,1].CurrentValue := -12.498303, [0,1].RangeMax := 50.0, [0,1].RangeMaxSave := 50.0, [0,1].RealCfg := 1, [0,1].EnableCfg := 1, [0,1].OverrideCfg := 1, [0,2].TagName := 'AI201A', [0,2].OutofRange := 1, [0,2].Address := 2, [0,2].RawMin := 5529, [0,2].RawMax := 27648, [0,2].RawLowLimit := 5253, [0,2].RawHighLimit := 27924, [0,2].FilterActual := 1.0, [0,2].ScaledMax := 100.0, [0,2].CurrentValue := -24.996607, [0,2].RangeMax := 100.0, [0,2].RangeMaxSave := 100.0, [0,2].RealCfg := 1, [0,2].EnableCfg := 1, [0,2].OverrideCfg := 1, [0,3].TagName := 'AI202', [0,3].OutofRange := 1, [0,3].Address := 3, [0,3].RawMin := 5529, [0,3].RawMax := 27648, [0,3].RawLowLimit := 5253, [0,3].RawHighLimit := 27924, [0,3].FilterActual := 1.0, [0,3].ScaledMax := 14.0, [0,3].CurrentValue := -3.499525, [0,3].RangeMax := 14.0, [0,3].RangeMaxSave := 14.0, [0,3].RealCfg := 1, [0,3].EnableCfg := 1,
        [0,3].OverrideCfg := 1, [0,4].TagName := 'TI201', [0,4].OutofRange := 1, [0,4].Address := 4, [0,4].RawMin := 5529, [0,4].RawMax := 27648, [0,4].RawLowLimit := 5253, [0,4].RawHighLimit := 27924, [0,4].FilterActual := 1.0, [0,4].ScaledMax := 100.0, [0,4].CurrentValue := -24.996607, [0,4].RangeMax := 100.0, [0,4].RangeMaxSave := 100.0, [0,4].RealCfg := 1, [0,4].EnableCfg := 1, [0,4].OverrideCfg := 1, [0,5].TagName := 'AI203', [0,5].OutofRange := 1, [0,5].Address := 5, [0,5].RawMin := 5529, [0,5].RawMax := 27648, [0,5].RawLowLimit := 5253, [0,5].RawHighLimit := 27924, [0,5].FilterActual := 1.0, [0,5].ScaledMax := 2.0, [0,5].CurrentValue := -0.49993217, [0,5].RangeMax := 2.0, [0,5].RangeMaxSave := 2.0, [0,5].RealCfg := 1, [0,5].EnableCfg := 1, [0,5].OverrideCfg := 1, [0,6].TagName := 'AI204', [0,6].OutofRange := 1, [0,6].Address := 6, [0,6].RawMin := 5529, [0,6].RawMax := 27648, [0,6].RawLowLimit := 5253, [0,6].RawHighLimit := 27924, [0,6].FilterActual := 1.0, [0,6].ScaledMax := 2.0, [0,6].CurrentValue := -0.49993217, [0,6].RangeMax := 2.0, [0,6].RangeMaxSave := 2.0, [0,6].RealCfg := 1, [0,6].EnableCfg := 1, [0,6].OverrideCfg := 1, [0,7].TagName := 'AI102', [0,7].OutofRange := 1, [0,7].Address := 7, [0,7].RawMin := 5529, [0,7].RawMax := 27648, [0,7].RawLowLimit := 5253, [0,7].RawHighLimit := 27924, [0,7].FilterActual := 1.0, [0,7].ScaledMax := 100.0, [0,7].CurrentValue := -24.996607, [0,7].RangeMax := 100.0, [0,7].RangeMaxSave := 100.0, [0,7].RealCfg := 1, [0,7].EnableCfg := 1,
        [0,7].OverrideCfg := 1, [0,8].TagName := 'AI103', [0,8].OutofRange := 1, [0,8].Address := 8, [0,8].RawMin := 5529, [0,8].RawMax := 27648, [0,8].RawLowLimit := 5253, [0,8].RawHighLimit := 27924, [0,8].FilterActual := 1.0, [0,8].ScaledMax := 14.0, [0,8].CurrentValue := -3.499525, [0,8].RangeMax := 14.0, [0,8].RangeMaxSave := 14.0, [0,8].RealCfg := 1, [0,8].EnableCfg := 1, [0,8].OverrideCfg := 1, [0,9].TagName := 'PI003', [0,9].OutofRange := 1, [0,9].Address := 9, [0,9].RawMin := 6553, [0,9].RawMax := 32767, [0,9].RawLowLimit := 6225, [0,9].RawHighLimit := 33095, [0,9].FilterActual := 1.0, [0,9].ScaledMax := 6.0, [0,9].CurrentValue := -1.4998856, [0,9].RangeMax := 6.0, [0,9].RangeMaxSave := 6.0, [0,9].RealCfg := 1, [0,9].EnableCfg := 1, [0,9].OverrideCfg := 1, [0,10].TagName := 'FI001', [0,10].Address := 10, [0,10].RawMin := 5529, [0,10].RawMax := 27648, [0,10].RawLowLimit := 5253, [0,10].RawHighLimit := 27924, [0,10].FilterActual := 1.0, [0,10].ScaledMax := 22.0, [0,10].RangeMax := 22.0, [0,10].RangeMaxSave := 22.0, [0,10].EnableCfg := 1, [0,10].OverrideCfg := 1, [0,11].TagName := 'PI001', [0,11].OutofRange := 1, [0,11].Address := 11, [0,11].RawMin := 6553, [0,11].RawMax := 32767, [0,11].RawLowLimit := 6225, [0,11].RawHighLimit := 33095, [0,11].FilterActual := 1.0, [0,11].ScaledMax := 6.0, [0,11].CurrentValue := -1.4998856, [0,11].RangeMax := 6.0, [0,11].RangeMaxSave := 6.0, [0,11].RealCfg := 1, [0,11].EnableCfg := 1, [0,11].OverrideCfg := 1, [0,12].TagName := 'FI002', [0,12].Address := 12,
        [0,12].RawMin := 5529, [0,12].RawMax := 27648, [0,12].RawLowLimit := 5253, [0,12].RawHighLimit := 27924, [0,12].FilterActual := 1.0, [0,12].ScaledMax := 22.0, [0,12].RangeMax := 22.0, [0,12].RangeMaxSave := 22.0, [0,12].EnableCfg := 1, [0,12].OverrideCfg := 1, [0,13].TagName := 'PI002', [0,13].OutofRange := 1, [0,13].Address := 13, [0,13].RawMin := 6553, [0,13].RawMax := 32767, [0,13].RawLowLimit := 6225, [0,13].RawHighLimit := 33095, [0,13].FilterActual := 1.0, [0,13].ScaledMax := 6.0, [0,13].CurrentValue := -1.4998856, [0,13].RangeMax := 6.0, [0,13].RangeMaxSave := 6.0, [0,13].RealCfg := 1, [0,13].EnableCfg := 1, [0,13].OverrideCfg := 1, [0,14].OutofRange := 1, [0,14].Address := 14, [0,14].RawMin := 5529, [0,14].RawMax := 27648, [0,14].RawLowLimit := 5253, [0,14].RawHighLimit := 27924, [0,14].FilterActual := 1.0, [0,14].ScaledMax := 14.0, [0,14].RangeMax := 14.0, [0,14].RangeMaxSave := 14.0, [0,14].RealCfg := 1, [0,14].OverrideCfg := 1, [0,15].OutofRange := 1, [0,15].Address := 15, [0,15].RawMin := 5529, [0,15].RawMax := 27648, [0,15].RawLowLimit := 5253, [0,15].RawHighLimit := 27924, [0,15].FilterActual := 1.0, [0,15].ScaledMax := 2.0, [0,15].CurrentValue := -0.49993217, [0,15].RangeMax := 2.0, [0,15].RangeMaxSave := 2.0, [0,15].RealCfg := 1, [0,15].OverrideCfg := 1, [0,16].OutofRange := 1, [0,16].Address := 16, [0,16].RawMin := 5529, [0,16].RawMax := 27648, [0,16].RawLowLimit := 5253, [0,16].RawHighLimit := 27924, [0,16].FilterActual := 1.0, [0,16].ScaledMax := 2.0, [0,16].CurrentValue := -0.49993217, [0,16].RangeMax := 2.0,
        [0,16].RangeMaxSave := 2.0, [0,16].RealCfg := 1, [0,16].OverrideCfg := 1, [0,17].OutofRange := 1, [0,17].Address := 17, [0,17].RawMin := 5529, [0,17].RawMax := 27648, [0,17].RawLowLimit := 5253, [0,17].RawHighLimit := 27924, [0,17].FilterActual := 1.0, [0,17].ScaledMin := -1.0, [0,17].ScaledMax := 5.0, [0,17].CurrentValue := -2.4997964, [0,17].RangeMin := -1.0, [0,17].RangeMax := 5.0, [0,17].RangeMinSave := -1.0, [0,17].RangeMaxSave := 5.0, [0,17].RealCfg := 1, [0,17].OverrideCfg := 1, [0,18].OutofRange := 1, [0,18].Address := 18, [0,18].RawMin := 5529, [0,18].RawMax := 27648, [0,18].RawLowLimit := 5253, [0,18].RawHighLimit := 27924, [0,18].FilterActual := 1.0, [0,18].ScaledMin := -1.0, [0,18].ScaledMax := 5.0, [0,18].CurrentValue := -2.4997964, [0,18].RangeMin := -1.0, [0,18].RangeMax := 5.0, [0,18].RangeMinSave := -1.0, [0,18].RangeMaxSave := 5.0, [0,18].RealCfg := 1, [0,18].OverrideCfg := 1, [0,19].OutofRange := 1, [0,19].Address := 19, [0,19].RawMin := 5529, [0,19].RawMax := 27648, [0,19].RawLowLimit := 5253, [0,19].RawHighLimit := 27924, [0,19].FilterActual := 1.0, [0,19].ScaledMin := -1.0, [0,19].ScaledMax := 5.0, [0,19].CurrentValue := -2.4997964, [0,19].RangeMin := -1.0, [0,19].RangeMax := 5.0, [0,19].RangeMinSave := -1.0, [0,19].RangeMaxSave := 5.0, [0,19].RealCfg := 1, [0,19].OverrideCfg := 1, [0,20].OutofRange := 1, [0,20].Address := 20, [0,20].RawMin := 5529, [0,20].RawMax := 27648, [0,20].RawLowLimit := 5253, [0,20].RawHighLimit := 27924, [0,20].FilterActual := 1.0, [0,20].ScaledMax := 100.0, [0,20].CurrentValue := -24.996607,
        [0,20].RangeMax := 100.0, [0,20].RangeMaxSave := 100.0, [0,20].RealCfg := 1, [0,20].OverrideCfg := 1, [0,21].OutofRange := 1, [0,21].Address := 21, [0,21].RawMin := 5529, [0,21].RawMax := 27648, [0,21].RawLowLimit := 5253, [0,21].RawHighLimit := 27924, [0,21].FilterActual := 1.0, [0,21].ScaledMax := 100.0, [0,21].CurrentValue := -24.996607, [0,21].RangeMax := 100.0, [0,21].RangeMaxSave := 100.0, [0,21].RealCfg := 1, [0,21].OverrideCfg := 1, [0,22].TagName := 'SPARE', [0,22].Address := 22, [0,22].RawMin := 5529, [0,22].RawMax := 27648, [0,22].RealCfg := 1, [0,22].OverrideCfg := 1, [0,23].TagName := 'SPARE', [0,23].Address := 23, [0,23].RawMin := 5529, [0,23].RawMax := 27648, [0,23].RealCfg := 1, [0,23].OverrideCfg := 1, [0,24].TagName := 'SPARE', [0,24].Address := 24, [0,24].RawMin := 5529, [0,24].RawMax := 27648, [0,24].RealCfg := 1, [0,24].OverrideCfg := 1, [0,25].TagName := 'SPARE', [0,25].Address := 25, [0,25].RawMin := 5529, [0,25].RawMax := 27648, [0,25].RealCfg := 1, [0,25].OverrideCfg := 1, [0,26].TagName := 'SPARE', [0,26].Address := 26, [0,26].RawMin := 5529, [0,26].RawMax := 27648, [0,26].RealCfg := 1, [0,26].OverrideCfg := 1, [0,27].TagName := 'SPARE', [0,27].Address := 27, [0,27].RawMin := 5529, [0,27].RawMax := 27648, [0,27].RealCfg := 1, [0,27].OverrideCfg := 1, [0,28].TagName := 'AI#1', [0,28].OutofRange := 1, [0,28].Address := 28, [0,28].RawMin := 6553, [0,28].RawMax := 32767, [0,28].RawLowLimit := 6225, [0,28].RawHighLimit := 33095,
        [0,28].FilterActual := 1.0, [0,28].ScaledMax := 100.0, [0,28].CurrentValue := -24.998093, [0,28].RangeMax := 100.0, [0,28].RangeMaxSave := 100.0, [0,28].RealCfg := 1, [0,28].EnableCfg := 1, [0,28].OverrideCfg := 1, [0,29].TagName := 'AI#2', [0,29].OutofRange := 1, [0,29].Address := 29, [0,29].RawMin := 6553, [0,29].RawMax := 32767, [0,29].RawLowLimit := 6225, [0,29].RawHighLimit := 33095, [0,29].FilterActual := 1.0, [0,29].ScaledMax := 100.0, [0,29].CurrentValue := -24.998093, [0,29].RangeMax := 100.0, [0,29].RangeMaxSave := 100.0, [0,29].RealCfg := 1, [0,29].EnableCfg := 1, [0,29].OverrideCfg := 1, [0,30].TagName := 'AI#3', [0,30].OutofRange := 1, [0,30].Address := 30, [0,30].RawMin := 6553, [0,30].RawMax := 32767, [0,30].RawValue := 49, [0,30].RawLowLimit := 6225, [0,30].RawHighLimit := 33095, [0,30].FilteredRaw := 49, [0,30].FilterActual := 1.0, [0,30].ScaledMax := 100.0, [0,30].CurrentValue := -24.811169, [0,30].RangeMax := 100.0, [0,30].RangeMaxSave := 100.0, [0,30].RealCfg := 1, [0,30].EnableCfg := 1, [0,30].OverrideCfg := 1, [0,31].TagName := 'AI#4', [0,31].OutofRange := 1, [0,31].Address := 31, [0,31].RawMin := 6553, [0,31].RawMax := 32767, [0,31].RawValue := 48, [0,31].RawLowLimit := 6225, [0,31].RawHighLimit := 33095, [0,31].FilteredRaw := 48, [0,31].FilterActual := 1.0, [0,31].ScaledMax := 100.0, [0,31].CurrentValue := -24.814985, [0,31].RangeMax := 100.0, [0,31].RangeMaxSave := 100.0, [0,31].RealCfg := 1, [0,31].EnableCfg := 1, [0,31].OverrideCfg := 1, [0,40].TagName := 'FI003', [0,40].Address := 40, [0,40].RawMin := 5529,
        [0,40].RawMax := 27648, [0,40].RawLowLimit := 5253, [0,40].RawHighLimit := 27924, [0,40].FilterActual := 1.0, [0,40].ScaledMax := 44.0, [0,40].RangeMax := 44.0, [0,40].RangeMaxSave := 44.0, [0,40].EnableCfg := 1, [0,40].OverrideCfg := 1, [0,41].TagName := 'LV003', [0,41].Address := 41, [0,41].RawMin := 6553, [0,41].RawMax := 32767, [0,41].RawLowLimit := 6225, [0,41].RawHighLimit := 33095, [0,41].FilterActual := 1.0, [0,41].ScaledMax := 9999.0, [0,41].RangeMax := 9999.0, [0,41].RangeMaxSave := 9999.0, [0,41].EnableCfg := 1, [0,41].OverrideCfg := 1, [0,42].TagName := 'LV001', [0,42].Address := 42, [0,42].RawMin := 6553, [0,42].RawMax := 32767, [0,42].RawLowLimit := 6225, [0,42].RawHighLimit := 33095, [0,42].FilterActual := 1.0, [0,42].ScaledMax := 9999.0, [0,42].RangeMax := 9999.0, [0,42].RangeMaxSave := 9999.0, [0,42].EnableCfg := 1, [0,42].OverrideCfg := 1, [0,43].TagName := 'LV002', [0,43].Address := 43, [0,43].RawMin := 6553, [0,43].RawMax := 32767, [0,43].RawLowLimit := 6225, [0,43].RawHighLimit := 33095, [0,43].FilterActual := 1.0, [0,43].ScaledMax := 9999.0, [0,43].RangeMax := 9999.0, [0,43].RangeMaxSave := 9999.0, [0,43].EnableCfg := 1, [0,43].OverrideCfg := 1, [0,44].Address := 44, [0,44].RawMin := 6553, [0,44].RawMax := 32767, [0,44].RawLowLimit := 6225, [0,44].RawHighLimit := 33095, [0,44].FilterActual := 1.0, [0,44].ScaledMax := 99999.0, [0,44].RangeMax := 99999.0, [0,44].RangeMaxSave := 99999.0, [0,45].Address := 42, [0,45].RawMin := 6553, [0,45].RawMax := 32767, [0,45].RawLowLimit := 6225, [0,45].RawHighLimit := 33095, [0,45].FilterActual := 1.0,
        [0,45].ScaledMin := -1.0, [0,45].ScaledMax := 5.0, [0,45].RangeMin := -1.0, [0,45].RangeMax := 5.0, [0,45].RangeMinSave := -1.0, [0,45].RangeMaxSave := 5.0, [0,45].OverrideCfg := 1, [1,0].TagName := 'WI101', [1,0].RawMax := 99999, [1,0].RawLowLimit := -1000, [1,0].RawHighLimit := 100999, [1,0].FilterActual := 1.0, [1,0].ScaledMax := 9999.9, [1,0].RangeMax := 600.0, [1,0].RangeMaxSave := 600.0, [1,0].EnableCfg := 1, [1,0].OverrideCfg := 1, [1,0].EGU := 'kg', [1,1].TagName := 'WI102', [1,1].OutofRange := 1, [1,1].Address := 1, [1,1].RawMin := 6553, [1,1].RawMax := 32767, [1,1].RawValue := 1, [1,1].RawLowLimit := 6225, [1,1].RawHighLimit := 33095, [1,1].FilterActual := 1.0, [1,1].ScaledMax := 50.0, [1,1].CurrentValue := -12.498811, [1,1].RangeMax := 50.0, [1,1].RangeMaxSave := 50.0, [1,1].OverrideCfg := 1, [1,2].TagName := 'FI101', [1,2].Address := 2, [1,2].RawMin := 6553, [1,2].RawMax := 32767, [1,2].RawValue := 6574, [1,2].RawLowLimit := 6225, [1,2].RawHighLimit := 33095, [1,2].FilteredRaw := 6574, [1,2].FilterActual := 1.0, [1,2].ScaledMax := 15.0, [1,2].CurrentValue := 0.01201648, [1,2].RangeMax := 15.0, [1,2].RangeMaxSave := 15.0, [1,2].RealCfg := 1, [1,2].EnableCfg := 1, [1,2].OverrideCfg := 1, [1,2].EGU := 'Lpm', [1,3].TagName := 'PCV001', [1,3].Address := 3, [1,3].RawMin := 6553, [1,3].RawMax := 32767, [1,3].RawValue := 23416, [1,3].RawLowLimit := 6225, [1,3].RawHighLimit := 33095, [1,3].FilteredRaw := 23416, [1,3].FilterActual := 1.0, [1,3].ScaledMax := 100.0, [1,3].CurrentValue := 101.99314,
        [1,3].RangeMax := 100.0, [1,3].RangeMaxSave := 100.0, [1,3].EnableCfg := 1, [1,3].EGU := '%Clo', [1,4].TagName := 'PCV101', [1,4].Address := 4, [1,4].RawMin := 6553, [1,4].RawMax := 32767, [1,4].RawValue := 21167, [1,4].RawLowLimit := 6225, [1,4].RawHighLimit := 33095, [1,4].FilteredRaw := 21167, [1,4].FilterActual := 1.0, [1,4].ScaledMax := 100.0, [1,4].CurrentValue := 38.696636, [1,4].RangeMax := 100.0, [1,4].RangeMaxSave := 100.0, [1,4].EnableCfg := 1, [1,4].EGU := '%Opn', [1,5].TagName := 'PI001', [1,5].Address := 5, [1,5].RawMin := 6553, [1,5].RawMax := 32767, [1,5].RawValue := 6505, [1,5].RawLowLimit := 6225, [1,5].RawHighLimit := 33095, [1,5].FilteredRaw := 6505, [1,5].FilterActual := 1.0, [1,5].ScaledMax := 6.0, [1,5].CurrentValue := -0.010986496, [1,5].RangeMax := 6.0, [1,5].RangeMaxSave := 6.0, [1,5].RealCfg := 1, [1,5].EnableCfg := 1, [1,5].OverrideCfg := 1, [1,5].EGU := 'bar', [1,6].TagName := 'PI002', [1,6].Address := 6, [1,6].RawMin := 6553, [1,6].RawMax := 32767, [1,6].RawValue := 6381, [1,6].RawLowLimit := 6225, [1,6].RawHighLimit := 33095, [1,6].FilterUser := 50, [1,6].FilteredRaw := 6386, [1,6].FilterActual := 0.5, [1,6].ScaledMax := 6.0, [1,6].CurrentValue := -0.03822385, [1,6].RangeMax := 6.0, [1,6].RangeMaxSave := 6.0, [1,6].RealCfg := 1, [1,6].EnableCfg := 1, [1,6].OverrideCfg := 1, [1,6].EGU := 'bar', [1,7].TagName := 'PI101', [1,7].Address := 7, [1,7].RawMin := 6553, [1,7].RawMax := 32767, [1,7].RawValue := 6486, [1,7].RawLowLimit := 6225,
        [1,7].RawHighLimit := 33095, [1,7].FilteredRaw := 6486, [1,7].FilterActual := 1.0, [1,7].ScaledMax := 6.0, [1,7].CurrentValue := -0.015335317, [1,7].RangeMax := 6.0, [1,7].RangeMaxSave := 6.0, [1,7].RealCfg := 1, [1,7].EnableCfg := 1, [1,7].OverrideCfg := 1, [1,7].EGU := 'bar', [1,8].TagName := 'PI401', [1,8].Address := 8, [1,8].RawMin := 6553, [1,8].RawMax := 32767, [1,8].RawValue := 6616, [1,8].RawLowLimit := 6225, [1,8].RawHighLimit := 33095, [1,8].FilteredRaw := 6616, [1,8].FilterActual := 1.0, [1,8].ScaledMax := 6.0, [1,8].CurrentValue := 0.014419775, [1,8].RangeMax := 6.0, [1,8].RangeMaxSave := 6.0, [1,8].RealCfg := 1, [1,8].EnableCfg := 1, [1,8].OverrideCfg := 1, [1,8].EGU := 'bar', [1,9].TagName := 'AI104', [1,9].OutofRange := 1, [1,9].Address := 9, [1,9].RawMin := 6553, [1,9].RawMax := 32767, [1,9].RawLowLimit := 6225, [1,9].RawHighLimit := 33095, [1,9].FilterActual := 1.0, [1,9].ScaledMax := 14.0, [1,9].RangeMax := 14.0, [1,9].RangeMaxSave := 14.0, [1,9].RealCfg := 1, [1,9].OverrideCfg := 1, [1,9].EGU := 'pH', [1,10].TagName := 'AI101', [1,10].Address := 10, [1,10].RawMin := 6553, [1,10].RawMax := 32767, [1,10].RawValue := 6558, [1,10].RawLowLimit := 6225, [1,10].RawHighLimit := 33095, [1,10].FilteredRaw := 6558, [1,10].FilterActual := 1.0, [1,10].ScaledMax := 100.0, [1,10].CurrentValue := 0.019073777, [1,10].RangeMax := 100.0, [1,10].RangeMaxSave := 100.0, [1,10].RealCfg := 1, [1,10].EnableCfg := 1, [1,10].OverrideCfg := 1, [1,10].EGU := '$B5S/cm', [1,11].TagName := 'AI102',
        [1,11].Address := 11, [1,11].RawMin := 6553, [1,11].RawMax := 32767, [1,11].RawValue := 6576, [1,11].RawLowLimit := 6225, [1,11].RawHighLimit := 33095, [1,11].FilteredRaw := 6576, [1,11].FilterActual := 1.0, [1,11].ScaledMax := 2.0, [1,11].CurrentValue := 0.0017547875, [1,11].RangeMax := 2.0, [1,11].RangeMaxSave := 2.0, [1,11].RealCfg := 1, [1,11].EnableCfg := 1, [1,11].OverrideCfg := 1, [1,11].EGU := 'AU', [1,12].TagName := 'AI103', [1,12].Address := 12, [1,12].RawMin := 6553, [1,12].RawMax := 32767, [1,12].RawValue := 6600, [1,12].RawLowLimit := 6225, [1,12].RawHighLimit := 33095, [1,12].FilteredRaw := 6600, [1,12].FilterActual := 1.0, [1,12].ScaledMax := 2.0, [1,12].CurrentValue := 0.0035858701, [1,12].RangeMax := 2.0, [1,12].RangeMaxSave := 2.0, [1,12].RealCfg := 1, [1,12].EnableCfg := 1, [1,12].OverrideCfg := 1, [1,12].EGU := 'AU', [1,13].TagName := 'TI001', [1,13].Address := 13, [1,13].RawMin := 6553, [1,13].RawMax := 32767, [1,13].RawValue := 17260, [1,13].RawLowLimit := 6225, [1,13].RawHighLimit := 33095, [1,13].FilteredRaw := 17260, [1,13].FilterActual := 1.0, [1,13].ScaledMax := 55.0, [1,13].CurrentValue := 22.464523, [1,13].RangeMax := 55.0, [1,13].RangeMaxSave := 55.0, [1,13].RealCfg := 1, [1,13].EnableCfg := 1, [1,13].OverrideCfg := 1, [1,13].EGU := '$B0C', [1,14].TagName := 'MIX001', [1,14].Address := 14, [1,14].RawMax := 16384, [1,14].RawValue := 42, [1,14].RawLowLimit := -164, [1,14].RawHighLimit := 16548, [1,14].FilteredRaw := 42, [1,14].FilterActual := 1.0, [1,14].ScaledMax := 100.0, [1,14].CurrentValue := 0.25634766,
        [1,14].RangeMax := 100.0, [1,14].RangeMaxSave := 100.0, [1,14].RealCfg := 1, [1,14].EnableCfg := 1, [1,14].EGU := '%', [1,15].TagName := 'WI001', [1,15].Address := 15, [1,15].RawMax := 99999, [1,15].RawValue := -16, [1,15].RawLowLimit := -1000, [1,15].RawHighLimit := 100999, [1,15].FilteredRaw := -16, [1,15].FilterActual := 1.0, [1,15].ScaledMax := 999.99, [1,15].CurrentValue := -0.16, [1,15].EnableCfg := 1, [1,15].OverrideCfg := 1, [1,16].TagName := 'WI101', [1,16].OutofRange := 1, [1,16].Address := 16, [1,16].RawMin := 5529, [1,16].RawMax := 27648, [1,16].RawLowLimit := 5253, [1,16].RawHighLimit := 27924, [1,16].FilterActual := 1.0, [1,16].ScaledMax := 2.0, [1,16].RangeMax := 2.0, [1,16].RangeMaxSave := 2.0, [1,16].RealCfg := 1, [1,16].OverrideCfg := 1, [1,17].TagName := 'FI003', [1,17].OutofRange := 1, [1,17].Address := 17, [1,17].RawMin := 6553, [1,17].RawMax := 32767, [1,17].RawLowLimit := 5253, [1,17].RawHighLimit := 27924, [1,17].FilterActual := 1.0, [1,17].ScaledMax := 15.0, [1,17].RangeMax := 15.0, [1,17].RangeMaxSave := 15.0, [1,17].RealCfg := 1, [1,17].OverrideCfg := 1, [1,18].OutofRange := 1, [1,18].Address := 18, [1,18].RawMin := 5529, [1,18].RawMax := 27648, [1,18].RawLowLimit := 5253, [1,18].RawHighLimit := 27924, [1,18].FilterActual := 1.0, [1,18].ScaledMin := -1.0, [1,18].ScaledMax := 5.0, [1,18].RangeMin := -1.0, [1,18].RangeMax := 5.0, [1,18].RangeMinSave := -1.0, [1,18].RangeMaxSave := 5.0, [1,18].RealCfg := 1, [1,18].OverrideCfg := 1, [1,19].OutofRange := 1, [1,19].Address := 19,
        [1,19].RawMin := 5529, [1,19].RawMax := 27648, [1,19].RawLowLimit := 5253, [1,19].RawHighLimit := 27924, [1,19].FilterActual := 1.0, [1,19].ScaledMin := -1.0, [1,19].ScaledMax := 5.0, [1,19].RangeMin := -1.0, [1,19].RangeMax := 5.0, [1,19].RangeMinSave := -1.0, [1,19].RangeMaxSave := 5.0, [1,19].RealCfg := 1, [1,19].OverrideCfg := 1, [1,20].OutofRange := 1, [1,20].Address := 20, [1,20].RawMin := 5529, [1,20].RawMax := 27648, [1,20].RawLowLimit := 5253, [1,20].RawHighLimit := 27924, [1,20].FilterActual := 1.0, [1,20].ScaledMax := 100.0, [1,20].RangeMax := 100.0, [1,20].RangeMaxSave := 100.0, [1,20].RealCfg := 1, [1,20].OverrideCfg := 1, [1,21].OutofRange := 1, [1,21].Address := 21, [1,21].RawMin := 5529, [1,21].RawMax := 27648, [1,21].RawLowLimit := 5253, [1,21].RawHighLimit := 27924, [1,21].FilterActual := 1.0, [1,21].ScaledMax := 100.0, [1,21].RangeMax := 100.0, [1,21].RangeMaxSave := 100.0, [1,21].RealCfg := 1, [1,21].OverrideCfg := 1, [1,22].TagName := 'SPARE', [1,22].Address := 22, [1,22].RawMin := 5529, [1,22].RawMax := 27648, [1,22].RealCfg := 1, [1,22].OverrideCfg := 1, [1,23].TagName := 'SPARE', [1,23].Address := 23, [1,23].RawMin := 5529, [1,23].RawMax := 27648, [1,23].RealCfg := 1, [1,23].OverrideCfg := 1, [1,24].TagName := 'SPARE', [1,24].Address := 24, [1,24].RawMin := 5529, [1,24].RawMax := 27648, [1,24].RealCfg := 1, [1,24].OverrideCfg := 1, [1,25].TagName := 'SPARE', [1,25].Address := 25, [1,25].RawMin := 5529, [1,25].RawMax := 27648, [1,25].RealCfg := 1,
        [1,25].OverrideCfg := 1, [1,26].TagName := 'SPARE', [1,26].Address := 26, [1,26].RawMin := 5529, [1,26].RawMax := 27648, [1,26].RealCfg := 1, [1,26].OverrideCfg := 1, [1,27].TagName := 'SPARE', [1,27].Address := 27, [1,27].RawMin := 5529, [1,27].RawMax := 27648, [1,27].RealCfg := 1, [1,27].OverrideCfg := 1, [1,28].OutofRange := 1, [1,28].Address := 28, [1,28].RawMin := 6553, [1,28].RawMax := 32767, [1,28].RawLowLimit := 6225, [1,28].RawHighLimit := 33095, [1,28].FilterActual := 1.0, [1,28].ScaledMax := 100.0, [1,28].CurrentValue := -24.998093, [1,28].RangeMax := 100.0, [1,28].RangeMaxSave := 100.0, [1,28].RealCfg := 1, [1,28].OverrideCfg := 1, [1,29].OutofRange := 1, [1,29].Address := 29, [1,29].RawMin := 6553, [1,29].RawMax := 32767, [1,29].RawLowLimit := 6225, [1,29].RawHighLimit := 33095, [1,29].FilterActual := 1.0, [1,29].ScaledMax := 100.0, [1,29].CurrentValue := -24.998093, [1,29].RangeMax := 100.0, [1,29].RangeMaxSave := 100.0, [1,29].RealCfg := 1, [1,29].OverrideCfg := 1, [1,30].OutofRange := 1, [1,30].Address := 30, [1,30].RawMin := 6553, [1,30].RawMax := 32767, [1,30].RawLowLimit := 6225, [1,30].RawHighLimit := 33095, [1,30].FilterActual := 1.0, [1,30].ScaledMax := 100.0, [1,30].CurrentValue := -24.998093, [1,30].RangeMax := 100.0, [1,30].RangeMaxSave := 100.0, [1,30].RealCfg := 1, [1,30].OverrideCfg := 1, [1,31].OutofRange := 1, [1,31].Address := 31, [1,31].RawMin := 6553, [1,31].RawMax := 32767, [1,31].RawLowLimit := 6225, [1,31].RawHighLimit := 33095, [1,31].FilterActual := 1.0, [1,31].ScaledMax := 100.0,
        [1,31].CurrentValue := -24.998093, [1,31].RangeMax := 100.0, [1,31].RangeMaxSave := 100.0, [1,31].RealCfg := 1, [1,31].OverrideCfg := 1, [1,40].TagName := 'DP', [1,40].Address := 40, [1,40].RawMin := 6553, [1,40].RawMax := 32767, [1,40].RawLowLimit := 6225, [1,40].RawHighLimit := 33095, [1,40].FilterActual := 1.0, [1,40].ScaledMax := 6.0, [1,40].CurrentValue := 0.026092928, [1,40].RangeMax := 6.0, [1,40].RangeMaxSave := 6.0, [1,40].EnableCfg := 1, [1,40].OverrideCfg := 1, [1,40].EGU := 'bar', [1,41].TagName := 'TMP', [1,41].Address := 41, [1,41].RawMin := 6553, [1,41].RawMax := 32767, [1,41].RawLowLimit := 6225, [1,41].RawHighLimit := 33095, [1,41].FilterActual := 1.0, [1,41].ScaledMax := 6.0, [1,41].CurrentValue := -0.009384299, [1,41].RangeMax := 6.0, [1,41].RangeMaxSave := 6.0, [1,41].EnableCfg := 1, [1,41].OverrideCfg := 1, [1,41].EGU := 'bar', [1,42].TagName := 'FI001', [1,42].Address := 42, [1,42].RawMin := 6553, [1,42].RawMax := 32767, [1,42].RawLowLimit := 6225, [1,42].RawHighLimit := 33095, [1,42].FilterActual := 1.0, [1,42].ScaledMax := 25.0, [1,42].RangeMax := 25.0, [1,42].RangeMaxSave := 25.0, [1,42].EnableCfg := 1, [1,42].OverrideCfg := 1, [1,42].EGU := 'Lpm', [1,43].TagName := 'FI401', [1,43].Address := 43, [1,43].RawMin := 6553, [1,43].RawMax := 32767, [1,43].RawLowLimit := 6225, [1,43].RawHighLimit := 33095, [1,43].FilterActual := 1.0, [1,43].ScaledMax := 25.0, [1,43].RangeMax := 25.0, [1,43].RangeMaxSave := 25.0, [1,43].EnableCfg := 1, [1,43].OverrideCfg := 1, [1,43].EGU := 'Lpm', [1,44].TagName := 'LI001',
        [1,44].Address := 44, [1,44].RawMin := 6553, [1,44].RawMax := 32767, [1,44].RawLowLimit := 6225, [1,44].RawHighLimit := 33095, [1,44].FilterActual := 1.0, [1,44].ScaledMax := 50.0, [1,44].CurrentValue := -0.16, [1,44].RangeMax := 50.0, [1,44].RangeMaxSave := 50.0, [1,44].EnableCfg := 1, [1,44].OverrideCfg := 1, [1,45].TagName := 'NWP', [1,45].Address := 45, [1,45].RawMin := 6553, [1,45].RawMax := 32767, [1,45].RawLowLimit := 6225, [1,45].RawHighLimit := 33095, [1,45].FilterActual := 1.0, [1,45].ScaledMax := 999.0, [1,45].CurrentValue := -81.47681, [1,45].RangeMax := 999.0, [1,45].RangeMaxSave := 999.0, [1,45].EnableCfg := 1, [1,45].EGU := 'Lm2h/', [1,46].TagName := 'PERM', [1,46].Address := 46, [1,46].RawMin := 6553, [1,46].RawMax := 32767, [1,46].RawLowLimit := 6225, [1,46].RawHighLimit := 33095, [1,46].FilterActual := 1.0, [1,46].ScaledMax := 999.0, [1,46].CurrentValue := -76.82927, [1,46].RangeMax := 999.0, [1,46].RangeMaxSave := 999.0, [1,46].EnableCfg := 1, [1,46].EGU := 'Lm2h/', [2,0].TagName := 'WI101', [2,0].RawMax := 99999, [2,0].RawLowLimit := -1000, [2,0].RawHighLimit := 100999, [2,0].FilterActual := 1.0, [2,0].ScaledMax := 9999.9, [2,0].RangeMax := 1500.0, [2,0].RangeMaxSave := 1500.0, [2,0].EnableCfg := 1, [2,0].OverrideCfg := 1, [2,0].EGU := 'kg', [2,1].TagName := 'WI102', [2,1].OutofRange := 1, [2,1].Address := 1, [2,1].RawMin := 6553, [2,1].RawMax := 32767, [2,1].RawLowLimit := 6225, [2,1].RawHighLimit := 33095, [2,1].FilterActual := 1.0, [2,1].ScaledMax := 50.0, [2,1].CurrentValue := -12.499105, [2,1].RangeMax := 50.0,
        [2,1].RangeMaxSave := 50.0, [2,1].OverrideCfg := 1, [2,2].TagName := 'FI101', [2,2].OutofRange := 1, [2,2].Address := 2, [2,2].RawMin := 6553, [2,2].RawMax := 32767, [2,2].RawLowLimit := 6225, [2,2].RawHighLimit := 33095, [2,2].FilterActual := 1.0, [2,2].ScaledMax := 25.0, [2,2].CurrentValue := -6.249523, [2,2].RangeMax := 25.0, [2,2].RangeMaxSave := 25.0, [2,2].RealCfg := 1, [2,2].EnableCfg := 1, [2,2].OverrideCfg := 1, [2,2].EGU := 'Lpm', [2,3].TagName := 'PCV001', [2,3].OutofRange := 1, [2,3].Address := 3, [2,3].RawMin := 6553, [2,3].RawMax := 32767, [2,3].RawLowLimit := 6225, [2,3].RawHighLimit := 33095, [2,3].FilterActual := 1.0, [2,3].ScaledMax := 100.0, [2,3].CurrentValue := -280.52606, [2,3].RangeMax := 100.0, [2,3].RangeMaxSave := 100.0, [2,3].EnableCfg := 1, [2,3].EGU := '%Clo', [2,4].TagName := 'PCV101', [2,4].OutofRange := 1, [2,4].Address := 4, [2,4].RawMin := 6553, [2,4].RawMax := 32767, [2,4].RawLowLimit := 6225, [2,4].RawHighLimit := 33095, [2,4].FilterActual := 1.0, [2,4].ScaledMax := 100.0, [2,4].CurrentValue := 380.95084, [2,4].RangeMax := 100.0, [2,4].RangeMaxSave := 100.0, [2,4].EnableCfg := 1, [2,4].EGU := '%Opn', [2,5].TagName := 'PI001', [2,5].OutofRange := 1, [2,5].Address := 5, [2,5].RawMin := 6553, [2,5].RawMax := 32767, [2,5].RawLowLimit := 6225, [2,5].RawHighLimit := 33095, [2,5].FilterActual := 1.0, [2,5].ScaledMax := 6.0, [2,5].CurrentValue := -1.4998856, [2,5].RangeMax := 6.0, [2,5].RangeMaxSave := 6.0, [2,5].RealCfg := 1, [2,5].EnableCfg := 1,
        [2,5].OverrideCfg := 1, [2,5].EGU := 'bar', [2,6].TagName := 'PI002', [2,6].OutofRange := 1, [2,6].Address := 6, [2,6].RawMin := 6553, [2,6].RawMax := 32767, [2,6].RawLowLimit := 6225, [2,6].RawHighLimit := 33095, [2,6].FilterUser := 50, [2,6].FilterActual := 0.5, [2,6].ScaledMax := 6.0, [2,6].CurrentValue := -1.4998856, [2,6].RangeMax := 6.0, [2,6].RangeMaxSave := 6.0, [2,6].RealCfg := 1, [2,6].EnableCfg := 1, [2,6].OverrideCfg := 1, [2,6].EGU := 'bar', [2,7].TagName := 'PI101', [2,7].OutofRange := 1, [2,7].Address := 7, [2,7].RawMin := 6553, [2,7].RawMax := 32767, [2,7].RawLowLimit := 6225, [2,7].RawHighLimit := 33095, [2,7].FilterActual := 1.0, [2,7].ScaledMax := 6.0, [2,7].CurrentValue := -1.4998856, [2,7].RangeMax := 6.0, [2,7].RangeMaxSave := 6.0, [2,7].RealCfg := 1, [2,7].EnableCfg := 1, [2,7].OverrideCfg := 1, [2,7].EGU := 'bar', [2,8].TagName := 'PI401', [2,8].OutofRange := 1, [2,8].Address := 8, [2,8].RawMin := 6553, [2,8].RawMax := 32767, [2,8].RawLowLimit := 6225, [2,8].RawHighLimit := 33095, [2,8].FilterActual := 1.0, [2,8].ScaledMax := 6.0, [2,8].CurrentValue := -1.4998856, [2,8].RangeMax := 6.0, [2,8].RangeMaxSave := 6.0, [2,8].RealCfg := 1, [2,8].EnableCfg := 1, [2,8].OverrideCfg := 1, [2,8].EGU := 'bar', [2,9].TagName := 'AI104', [2,9].OutofRange := 1, [2,9].Address := 9, [2,9].RawMin := 6553, [2,9].RawMax := 32767, [2,9].RawLowLimit := 6225, [2,9].RawHighLimit := 33095, [2,9].FilterActual := 1.0, [2,9].ScaledMax := 14.0,
        [2,9].CurrentValue := -1.4998856, [2,9].RangeMax := 14.0, [2,9].RangeMaxSave := 14.0, [2,9].RealCfg := 1, [2,9].OverrideCfg := 1, [2,9].EGU := 'pH', [2,10].TagName := 'AI101', [2,10].OutofRange := 1, [2,10].Address := 10, [2,10].RawMin := 6553, [2,10].RawMax := 32767, [2,10].RawLowLimit := 6225, [2,10].RawHighLimit := 33095, [2,10].FilterActual := 1.0, [2,10].ScaledMax := 100.0, [2,10].CurrentValue := -24.998093, [2,10].RangeMax := 100.0, [2,10].RangeMaxSave := 100.0, [2,10].RealCfg := 1, [2,10].EnableCfg := 1, [2,10].OverrideCfg := 1, [2,10].EGU := '$B5S/cm', [2,11].TagName := 'AI102', [2,11].OutofRange := 1, [2,11].Address := 11, [2,11].RawMin := 6553, [2,11].RawMax := 32767, [2,11].RawLowLimit := 6225, [2,11].RawHighLimit := 33095, [2,11].FilterActual := 1.0, [2,11].ScaledMax := 2.0, [2,11].CurrentValue := -0.49996185, [2,11].RangeMax := 2.0, [2,11].RangeMaxSave := 2.0, [2,11].RealCfg := 1, [2,11].OverrideCfg := 1, [2,11].EGU := 'AU', [2,12].TagName := 'AI103', [2,12].OutofRange := 1, [2,12].Address := 12, [2,12].RawMin := 6553, [2,12].RawMax := 32767, [2,12].RawLowLimit := 6225, [2,12].RawHighLimit := 33095, [2,12].FilterActual := 1.0, [2,12].ScaledMax := 2.0, [2,12].CurrentValue := -0.49996185, [2,12].RangeMax := 2.0, [2,12].RangeMaxSave := 2.0, [2,12].RealCfg := 1, [2,12].OverrideCfg := 1, [2,12].EGU := 'AU', [2,13].TagName := 'TI001', [2,13].OutofRange := 1, [2,13].Address := 13, [2,13].RawMin := 6553, [2,13].RawMax := 32767, [2,13].RawLowLimit := 6225, [2,13].RawHighLimit := 33095, [2,13].FilterActual := 1.0,
        [2,13].ScaledMax := 55.0, [2,13].CurrentValue := -13.748952, [2,13].RangeMax := 55.0, [2,13].RangeMaxSave := 55.0, [2,13].RealCfg := 1, [2,13].EnableCfg := 1, [2,13].OverrideCfg := 1, [2,13].EGU := '$B0C', [2,14].TagName := 'MIX001', [2,14].Address := 14, [2,14].RawMax := 16384, [2,14].RawLowLimit := -164, [2,14].RawHighLimit := 16548, [2,14].FilterActual := 1.0, [2,14].ScaledMax := 100.0, [2,14].RangeMax := 100.0, [2,14].RangeMaxSave := 100.0, [2,14].RealCfg := 1, [2,14].EnableCfg := 1, [2,14].EGU := '%', [2,15].TagName := 'WI001', [2,15].Address := 15, [2,15].RawMax := 99999, [2,15].RawLowLimit := -1000, [2,15].RawHighLimit := 100999, [2,15].FilterActual := 1.0, [2,15].ScaledMax := 999.99, [2,15].EnableCfg := 1, [2,15].OverrideCfg := 1, [2,16].CurrentValue := -0.4999322, [2,17].CurrentValue := -2.499796, [2,18].CurrentValue := -2.499796, [2,19].CurrentValue := -2.499796, [2,20].CurrentValue := -24.99661, [2,21].CurrentValue := -24.99661, [2,22].TagName := 'SPARE', [2,23].TagName := 'SPARE', [2,24].TagName := 'SPARE', [2,25].TagName := 'SPARE', [2,26].TagName := 'SPARE', [2,27].TagName := 'SPARE', [2,28].TagName := 'AI#1', [2,28].Address := 28, [2,28].RawMin := 6553, [2,28].RawMax := 32767, [2,28].RawValue := 12544, [2,28].RawLowLimit := 6225, [2,28].RawHighLimit := 33095, [2,28].FilteredRaw := 12544, [2,28].FilterActual := 1.0, [2,28].ScaledMax := 100.0, [2,28].CurrentValue := 22.8542, [2,28].RangeMax := 100.0, [2,28].RangeMaxSave := 100.0, [2,28].RealCfg := 1, [2,28].OverrideCfg := 1, [2,29].TagName := 'AI#2', [2,29].Address := 29, [2,29].RawMin := 6553, [2,29].RawMax := 32767,
        [2,29].RawValue := 12288, [2,29].RawLowLimit := 6225, [2,29].RawHighLimit := 33095, [2,29].FilteredRaw := 12288, [2,29].FilterActual := 1.0, [2,29].ScaledMax := 100.0, [2,29].CurrentValue := 21.877623, [2,29].RangeMax := 100.0, [2,29].RangeMaxSave := 100.0, [2,29].RealCfg := 1, [2,29].OverrideCfg := 1, [2,30].TagName := 'AI#3', [2,30].Address := 30, [2,30].RawMin := 6553, [2,30].RawMax := 32767, [2,30].RawValue := 12288, [2,30].RawLowLimit := 6225, [2,30].RawHighLimit := 33095, [2,30].FilteredRaw := 12288, [2,30].FilterActual := 1.0, [2,30].ScaledMax := 100.0, [2,30].CurrentValue := 21.877623, [2,30].RangeMax := 100.0, [2,30].RangeMaxSave := 100.0, [2,30].RealCfg := 1, [2,30].OverrideCfg := 1, [2,31].TagName := 'AI#4', [2,31].Address := 31, [2,31].RawMin := 6553, [2,31].RawMax := 32767, [2,31].RawValue := 12288, [2,31].RawLowLimit := 6225, [2,31].RawHighLimit := 33095, [2,31].FilteredRaw := 12288, [2,31].FilterActual := 1.0, [2,31].ScaledMax := 100.0, [2,31].CurrentValue := 21.877623, [2,31].RangeMax := 100.0, [2,31].RangeMaxSave := 100.0, [2,31].RealCfg := 1, [2,31].OverrideCfg := 1, [2,40].TagName := 'DP', [2,40].Address := 40, [2,40].RawMin := 6553, [2,40].RawMax := 32767, [2,40].RawLowLimit := 6225, [2,40].RawHighLimit := 33095, [2,40].FilterActual := 1.0, [2,40].ScaledMax := 6.0, [2,40].RangeMax := 6.0, [2,40].RangeMaxSave := 6.0, [2,40].EnableCfg := 1, [2,40].OverrideCfg := 1, [2,40].EGU := 'bar', [2,41].TagName := 'TMP', [2,41].Address := 41, [2,41].RawMin := 6553, [2,41].RawMax := 32767, [2,41].RawLowLimit := 6225, [2,41].RawHighLimit := 33095,
        [2,41].FilterActual := 1.0, [2,41].ScaledMax := 6.0, [2,41].RangeMax := 6.0, [2,41].RangeMaxSave := 6.0, [2,41].EnableCfg := 1, [2,41].OverrideCfg := 1, [2,41].EGU := 'bar', [2,42].TagName := 'FI001', [2,42].Address := 42, [2,42].RawMin := 6553, [2,42].RawMax := 32767, [2,42].RawLowLimit := 6225, [2,42].RawHighLimit := 33095, [2,42].FilterActual := 1.0, [2,42].ScaledMax := 45.0, [2,42].RangeMax := 45.0, [2,42].RangeMaxSave := 45.0, [2,42].EnableCfg := 1, [2,42].OverrideCfg := 1, [2,42].EGU := 'Lpm', [2,43].TagName := 'FI401', [2,43].Address := 43, [2,43].RawMin := 6553, [2,43].RawMax := 32767, [2,43].RawLowLimit := 6225, [2,43].RawHighLimit := 33095, [2,43].FilterActual := 1.0, [2,43].ScaledMax := 25.0, [2,43].RangeMax := 25.0, [2,43].RangeMaxSave := 25.0, [2,43].EnableCfg := 1, [2,43].OverrideCfg := 1, [2,43].EGU := 'Lpm', [2,44].TagName := 'LI001', [2,44].Address := 44, [2,44].RawMin := 6553, [2,44].RawMax := 32767, [2,44].RawLowLimit := 6225, [2,44].RawHighLimit := 33095, [2,44].FilterActual := 1.0, [2,44].ScaledMax := 50.0, [2,44].RangeMax := 50.0, [2,44].RangeMaxSave := 50.0, [2,44].EnableCfg := 1, [2,44].OverrideCfg := 1, [2,45].TagName := 'NWP', [2,45].Address := 45, [2,45].RawMin := 6553, [2,45].RawMax := 32767, [2,45].RawLowLimit := 6225, [2,45].RawHighLimit := 33095, [2,45].FilterActual := 1.0, [2,45].ScaledMax := 999.0, [2,45].RangeMax := 999.0, [2,45].RangeMaxSave := 999.0, [2,45].EnableCfg := 1, [2,45].EGU := 'Lm2h/', [2,46].TagName := 'PERM', [2,46].Address := 46, [2,46].RawMin := 6553,
        [2,46].RawMax := 32767, [2,46].RawLowLimit := 6225, [2,46].RawHighLimit := 33095, [2,46].FilterActual := 1.0, [2,46].ScaledMax := 999.0, [2,46].RangeMax := 999.0, [2,46].RangeMaxSave := 999.0, [2,46].EnableCfg := 1, [2,46].EGU := 'Lm2h/', [3,0].OutofRange := 1, [3,0].RawMin := 6553, [3,0].RawMax := 32767, [3,0].RawLowLimit := 6225, [3,0].RawHighLimit := 33095, [3,0].FilterActual := 1.0, [3,0].RealCfg := 1, [3,0].EnableCfg := 1, [3,0].OverrideCfg := 1, [3,1].TagName := 'PI002', [3,1].TagDisplayName := 'PI002', [3,1].OutofRange := 1, [3,1].Address := 1, [3,1].RawMin := 5529, [3,1].RawMax := 27648, [3,1].RawLowLimit := 5253, [3,1].RawHighLimit := 27924, [3,1].FilterUser := 50, [3,1].FilterActual := 0.5, [3,1].ScaledMax := 6.0, [3,1].CurrentValue := -0.06111238, [3,1].RangeMax := 6.0, [3,1].RangeMaxSave := 6.0, [3,1].RealCfg := 1, [3,1].EnableCfg := 1, [3,1].OverrideCfg := 1, [3,1].Desc := 'Retentate Pressure', [3,1].EGU := 'bar', [3,2].TagName := 'PI101', [3,2].TagDisplayName := 'PI101', [3,2].OutofRange := 1, [3,2].Address := 2, [3,2].RawMin := 5529, [3,2].RawMax := 27648, [3,2].RawLowLimit := 5253, [3,2].RawHighLimit := 27924, [3,2].FilterUser := 50, [3,2].FilterActual := 0.5, [3,2].ScaledMax := 6.0, [3,2].CurrentValue := -0.03822385, [3,2].RangeMax := 6.0, [3,2].RangeMaxSave := 6.0, [3,2].RealCfg := 1, [3,2].EnableCfg := 1, [3,2].OverrideCfg := 1, [3,2].Desc := 'Filtrate Pressure', [3,2].EGU := 'bar', [3,3].TagName := 'PI006', [3,3].TagDisplayName := 'PI006', [3,3].OutofRange := 1, [3,3].Address := 3,
